(* IEC 61131-3 sources: daoli-st-library/DL_Device (part 19) *)

(* ---- FB_DL_DieCastCycleSupervise.st ---- *)
(*==============================================================================
  Component : FB_DL_DieCastCycleSupervise
  Category  : DL_Device
  Type      : FB
  Complexity: C4
  VERSION   : v1.0.0
  功能      : 压铸单循环监控与三级异常分级停机（黄记录 / 红判废 / 黑停机）
  开源溯源  : 道莅原创 clean-room 自研（无外部代码引用）｜License: MIT
  边界条件  : ① 压射曲线四点监控：慢速终点位置偏差（eSlowEndDev）、快射峰值速度（eFastVelLow）、
                 增压建立时间（eBuildSlow）、保压压力（eHoldLow）；四点各自独立判据与独立成因，
                 分级动作经 ApplyDefect 单点施加，禁共用枚举成员（R190）。
              ② 分级语义（写进契约）：黄 = 记录成因、本模继续；红 = 置 _bRejectMark 判废并单拍告警，
                 机械流程仍走到 eDone 才结算（废件必须被顶出取走，不得停在模内）；
                 黑 = 立即停机（超压 / 信号非有限 / 急停 / 安全门开），等 bReset 复位。
              ③ 判据限值配比约束（R100）：fSlowEndWarnMm ≤ fSlowEndTolMm、fFastVelWarnMps ≥ fFastVelMinMps、
                 fBuildWarnS ≤ fBuildMaxS、fHoldWarnMpa ≥ fHoldMinMpa；违反即组态非法（E2 黑前哨）。
              ④ 默认引脚组合自证（R114）：过程握手类（bClampClosed / bClampOpened / bEjectDone /
                 bPartTaken / bSprayDone / bRejectAck）默认 FALSE，默认组合无法推进任何相；使能类
                 （bEStopHealthy / bGuardClosed）默认 TRUE 与 bEnable 同族，断线由硬件安全回路保证。
              ⑤ 复位作用域（R311）：bReset 沿清 E2/E3 锁存 + 判废标记 + 分级 + 曲线锁存；bStop 只清 E2 与相位。
  状态机    : eIdle 待机 / eClampClose 合模 / eShotSlow 慢压射 / eShotFast 快压射 / eIntensify 增压 /
              eHold 保压 / eClampOpen 开模 / eEject 顶出 / eTakeOut 取件 / eSpray 喷涂 / eDone 结算拍 /
              eFault 停机待复位(E2) / eSafeStop 安全断能(E3)
  自检      : R1 零 GVL ｜ R2 零物理地址 ｜ R3 纯 IEC 61131-3 ｜ R4 非有限自反判 + 除法先判分母 ｜
              R6 CASE 含 ELSE ｜ R7 九 TON 两沿段 0 无条件刷新 ｜ R10 仅标准转换函数 ｜ R14 无属性件
==============================================================================*)
TYPE E_DL_DcsPhase :
(
    eIdle       := 0,   (* 待机：等启动沿 / Idle, waiting for start edge *)
    eClampClose := 10,  (* 合模：等合模到位 / Clamp closing *)
    eShotSlow   := 20,  (* 慢压射：到慢速终点 / Slow shot *)
    eShotFast   := 30,  (* 快压射：到快射终点 / Fast shot *)
    eIntensify  := 40,  (* 增压：建压到门限 / Intensification *)
    eHold       := 50,  (* 保压：保压到时 / Pressure hold *)
    eClampOpen  := 60,  (* 开模：等开模到位 / Clamp opening *)
    eEject      := 70,  (* 顶出：等顶出到位 / Ejecting *)
    eTakeOut    := 80,  (* 取件：等取件完成 / Take-out *)
    eSpray      := 90,  (* 喷涂：等喷涂完成 / Spraying *)
    eDone       := 100, (* 结算拍：模次与良率统计 / Settlement, one-scan *)
    eFault      := 120, (* 停机待复位（E2）/ Stop awaiting reset, E2 *)
    eSafeStop   := 130  (* 安全侧断能（E3）/ Safety energy cut, E3 *)
);
END_TYPE
TYPE E_DL_DcsCause :
(
    eNone       := 0,   (* 无异常 / No anomaly *)
    eSlowEndDev := 1,   (* 慢速终点位置偏差超限（红）/ Slow-shot end position deviation *)
    eFastVelLow := 2,   (* 快射速度偏低（黄或红）/ Fast-shot velocity low *)
    eBuildSlow  := 3,   (* 增压建立时间超限（黄或红）/ Intensification build too slow *)
    eHoldLow    := 4,   (* 保压压力偏低（黄或红）/ Hold pressure low *)
    ePressOver  := 5,   (* 压力超上限（黑）/ Over-pressure, black *)
    eSigBad     := 6,   (* 压力或位置信号非有限（黑）/ Non-finite signal, black *)
    eEStopOpen  := 7,   (* 急停回路断开（黑）/ E-stop open, black *)
    eGuardOpen  := 8,   (* 安全门未闭合（黑）/ Guard door open, black *)
    eClampTmo   := 9,   (* 合模或开模超时（黑）/ Clamp timeout, black *)
    eShotTmo    := 10,  (* 压射超时（黑）/ Shot timeout, black *)
    eBuildTmo   := 11,  (* 增压超时（黑）/ Intensify timeout, black *)
    eFastTmo    := 12,  (* 快射超时（黑）/ Fast-shot timeout, black *)
    eEjectTmo   := 13,  (* 顶出超时（黑）/ Eject timeout, black *)
    eTakeTmo    := 14,  (* 取件超时（黑）/ Take-out timeout, black *)
    eSprayTmo   := 15,  (* 喷涂超时（黑）/ Spray timeout, black *)
    eCfgBad     := 16,  (* 组态非法（E2）/ Illegal configuration, E2 *)
    ePhaseBad   := 17   (* 非法相位兜底（E2）/ Illegal phase fallback, E2 *)
);
END_TYPE
TYPE E_DL_DcsGrade :
(
    eOk     := 0,       (* 无异常：本模继续 / OK, continue *)
    eYellow := 1,       (* 黄：记录并继续，不置 bError / Yellow, recorded only *)
    eRed    := 2,       (* 红：本模判废并告警 / Red, part rejected with alarm *)
    eBlack  := 3        (* 黑：立即停机 / Black, immediate stop *)
);
END_TYPE

FUNCTION_BLOCK FB_DL_DieCastCycleSupervise
VAR_INPUT
    bStart          : BOOL := FALSE;    (* 启动沿（eIdle 入 eClampClose） [-] / Start rising edge *)
    bStop           : BOOL := FALSE;    (* 中止：回 eIdle 并清 E2 锁存 [-] / Abort, clears E2 only *)
    bReset          : BOOL := FALSE;    (* 复位沿：清全部锁存 + 曲线锁存（R311） [-] / Reset edge *)
    bRejectAck      : BOOL := FALSE;    (* 废模确认（只清告警标记，不推进相） [-] / Reject acknowledge *)
    bClampClosed    : BOOL := FALSE;    (* 合模到位（默认 FALSE 禁跳步） [-] / Clamp closed *)
    bClampOpened    : BOOL := FALSE;    (* 开模到位（默认 FALSE 禁跳步） [-] / Clamp opened *)
    bEjectDone      : BOOL := FALSE;    (* 顶出到位（默认 FALSE 禁跳步） [-] / Eject done *)
    bPartTaken      : BOOL := FALSE;    (* 取件完成（默认 FALSE 禁跳步） [-] / Part taken *)
    bSprayDone      : BOOL := FALSE;    (* 喷涂完成（默认 FALSE 禁跳步） [-] / Spray done *)
    bGuardClosed    : BOOL := TRUE;     (* 安全门闭合（使能类引脚，默认 TRUE） [-] / Guard door closed *)
    bEStopHealthy   : BOOL := TRUE;     (* 急停回路正常（使能类引脚，默认 TRUE） [-] / E-stop healthy *)
    fShotPosMm      : LREAL := 0.0;     (* 冲头实时位置（0 = 起始位） [mm] / Shot position [mm] *)
    fShotVelMps     : LREAL := 0.0;     (* 冲头实时速度 [m/s] / Shot velocity [m/s] *)
    fHoldPressMpa   : LREAL := 0.0;     (* 压射缸压力实测 [MPa] / Shot pressure [MPa] *)
    fSlowEndSetMm   : LREAL := 250.0;   (* 慢速终点设定位置，域 > 0 [mm] / Slow-end setpoint [mm] *)
    fShotEndMm      : LREAL := 320.0;   (* 快射终点位置，域 > fSlowEndSetMm [mm] / Fast-shot end [mm] *)
    fSlowEndWarnMm  : LREAL := 10.0;    (* 慢速终点偏差预警限（黄），域 >= 0 [mm] / Slow-end warn limit [mm] *)
    fSlowEndTolMm   : LREAL := 25.0;    (* 慢速终点偏差硬限（红），域 > 0 [mm] / Slow-end hard limit [mm] *)
    fFastVelMinMps  : LREAL := 2.5;     (* 快射速度硬下限（红），域 > 0 [m/s] / Fast velocity hard min [m/s] *)
    fFastVelWarnMps : LREAL := 3.0;     (* 快射速度预警下限（黄），域 > 0 [m/s] / Fast velocity warn min [m/s] *)
    fIntensifyMpa   : LREAL := 18.0;    (* 增压建立压力门限，域 > 0 [MPa] / Build threshold [MPa] *)
    fBuildWarnS     : LREAL := 0.08;    (* 增压建立时间预警限（黄），域 >= 0 [s] / Build warn limit [s] *)
    fBuildMaxS      : LREAL := 0.15;    (* 增压建立时间硬限（红），域 > 0 [s] / Build hard limit [s] *)
    fHoldMinMpa     : LREAL := 12.0;    (* 保压压力硬下限（红），域 > 0 [MPa] / Hold pressure hard min [MPa] *)
    fHoldWarnMpa    : LREAL := 14.0;    (* 保压压力预警下限（黄），域 > 0 [MPa] / Hold pressure warn min [MPa] *)
    fPressOverMpa   : LREAL := 30.0;    (* 压力超上限（黑断能），域 > 0 [MPa] / Over-pressure limit [MPa] *)
    atPhaseTmo      : ARRAY[0..8] OF TIME := [T#10S, T#5S, T#5S, T#5S, T#30S, T#10S, T#10S, T#15S, T#15S];   (* 超时窗 [ms]，下标 0..8 = 合模/慢射/快射/增压/保压/开模/顶出/取件/喷涂 / Phase windows [ms] *)
    fCycleSec       : LREAL := 0.0;     (* 扫描周期（<=0 用缺省 0.01s） [s] / Scan cycle [s] *)
END_VAR
VAR_OUTPUT
    eState          : E_DL_DcsPhase;    (* 当前相（HMI 诊断） [-] / Present phase *)
    eCause          : E_DL_DcsCause;    (* 成因（锁存回放，R189） [-] / Latched cause playback *)
    eGrade          : E_DL_DcsGrade;    (* 本模判据分级（黄/红/黑）；组态 E2 不改分级、由 bError 表达 [-] / Criterion grade, E2 config fault expressed by bError *)
    bError          : BOOL;             (* 故障标志（仅黑与 E2 置位，黄/红不置） [-] / Error flag *)
    bSafeCut        : BOOL;             (* 安全侧断能指令（黑常 TRUE 至复位） [-] / Safety energy cut *)
    bReject         : BOOL;             (* 本模判废标告警（红级置位，结算或确认后清） [-] / Reject alarm *)
    bDone           : BOOL;             (* 单拍结算脉冲 [-] / One-scan done pulse *)
    bShotActive     : BOOL;             (* 压射段指示（供 IO 层驱动压射阀） [-] / Shot indicator *)
    nShotCount      : UDINT;            (* 累计模次（饱和） [模] / Shot count, saturating *)
    nGoodCount      : UDINT;            (* 累计良品（饱和） [模] / Good part count *)
    fYieldPct       : LREAL;            (* 良率（无模次输出 0） [%] / Yield [%] *)
    fSlowEndLastMm  : LREAL;            (* 最近一模慢速终点实测 [mm] / Last slow-end position [mm] *)
    fFastVelLastMps : LREAL;            (* 最近一模快射峰值速度 [m/s] / Last peak velocity [m/s] *)
    fBuildLastS     : LREAL;            (* 最近一模增压建立时间 [s] / Last build time [s] *)
    fHoldLastMpa    : LREAL;            (* 最近一模保压压力 [MPa] / Last hold pressure [MPa] *)
END_VAR
VAR
    _ePhase      : E_DL_DcsPhase := E_DL_DcsPhase.eIdle;     (* 内部相（CASE 唯一写入目标） [-] / Internal phase *)
    _eCause      : E_DL_DcsCause := E_DL_DcsCause.eNone;     (* 成因锁存量 [-] / Latched cause *)
    _eGrade      : E_DL_DcsGrade := E_DL_DcsGrade.eOk;       (* 本模分级锁存量 [-] / Latched grade *)
    _bFault      : BOOL := FALSE;       (* E2 锁存位（解除 = bReset 沿或 bStop） [-] / E2 latch *)
    _bSafeLatch  : BOOL := FALSE;       (* E3 锁存位（解除 = bReset 沿且安全恢复） [-] / E3 latch *)
    _bFaultReq   : BOOL := FALSE;       (* 单拍 E2 请求（段 1 预清，段 6 落地） [-] / One-scan E2 request *)
    _bSafeReq    : BOOL := FALSE;       (* 单拍 E3 请求（段 1 预清，段 6 落地） [-] / One-scan E3 request *)
    _bDonePulse  : BOOL := FALSE;       (* 单拍结算标志（段 1 预清） [-] / One-scan done flag *)
    _bRejectMark : BOOL := FALSE;       (* 本模判废标记（红级置位，结算清零） [-] / Reject mark for this shot *)
    _bPressBad   : BOOL := FALSE;       (* 压力信号非有限当拍量 [-] / Pressure non-finite *)
    _bPosBad     : BOOL := FALSE;       (* 位置信号非有限当拍量 [-] / Position non-finite *)
    _bVelBad     : BOOL := FALSE;       (* 速度信号非有限当拍量 [-] / Velocity non-finite *)
    _bBuilt      : BOOL := FALSE;       (* 增压已建立（当拍判据） [-] / Intensification built *)
    _bCfgBad     : BOOL := FALSE;       (* 组态非法当拍量 [-] / Configuration bad *)
    _nIdxChk     : INT := 0;            (* 相窗遍历索引（循环变量） [-] / Loop index *)
    _fCy         : LREAL := 0.0;        (* 当拍有效周期 [s] / Effective cycle *)
    _fVelPeak    : LREAL := 0.0;        (* 快射峰值速度（入快射相清零） [m/s] / Fast-shot peak [m/s] *)
    _fBuildS     : LREAL := 0.0;        (* 增压建立时间累加（入增压相清零） [s] / Build time accumulator [s] *)
    _fSlowEndMm  : LREAL := 0.0;        (* 慢速终点位置锁存 [mm] / Slow-end position latch *)
    _fHoldMpa    : LREAL := 0.0;        (* 保压压力锁存 [MPa] / Hold pressure latch *)
    _nShot       : UDINT := 0;          (* 模次累计锁存（饱和） [模] / Shot count latch *)
    _nGood       : UDINT := 0;          (* 良品累计锁存（饱和） [模] / Good count latch *)
    tonClampClose: TON;                 (* 合模超时（段 0 无条件调用） / Clamp-close timeout *)
    tonShotSlow  : TON;                 (* 慢压射超时 / Slow-shot timeout *)
    tonShotFast  : TON;                 (* 快压射超时 / Fast-shot timeout *)
    tonIntensify : TON;                 (* 增压超时 / Intensify timeout *)
    tonHold      : TON;                 (* 保压计时与超时 / Hold timer *)
    tonClampOpen : TON;                 (* 开模超时 / Clamp-open timeout *)
    tonEject     : TON;                 (* 顶出超时 / Eject timeout *)
    tonTakeOut   : TON;                 (* 取件超时 / Take-out timeout *)
    tonSpray     : TON;                 (* 喷涂超时 / Spray timeout *)
    rtStart      : R_TRIG;              (* 启动沿（段 0 无条件调用） / Start edge *)
    rtReset      : R_TRIG;              (* 复位沿（段 0 无条件调用） / Reset edge *)
END_VAR
VAR CONSTANT
    DL_DCS_CYDEF   : LREAL := 0.01;         (* 缺省扫描周期 [s] / Default scan cycle [s] *)
    DL_DCS_CNTMAX  : UDINT := 4294967295;   (* 模次与良品计数饱和上限 [模] / Count ceiling *)
    DL_DCS_PCTOP   : LREAL := 100.0;        (* 良率百分比满量程 [%] / Yield full scale [%] *)
END_VAR

(*-----------------------------------------------------------------------------
  方法 GradeFault：单点判据分级（纯分类，不修改任何 FB 状态）
  契约：fValue 为「按变差方向已归一」的判据量（偏差取绝对值后传入）；
        bLowerWorse = TRUE 表示低于限值变差，FALSE 表示高于限值变差；
        fWarnLimit 必须落在「正常侧」，fHardLimit 落在「变差侧」（配比由组态闸保证）。
        非有限实测（NaN 自反 / Inf 差值自减）一律返回 eBlack：信号失效必须停机。
-----------------------------------------------------------------------------*)
METHOD PUBLIC GradeFault : E_DL_DcsGrade
VAR_INPUT
    fValue      : LREAL := 0.0;     (* 判据实测值（已按方向归一） [工程单位] / Measured criterion *)
    fWarnLimit  : LREAL := 0.0;     (* 预警限（黄级） [工程单位] / Warning limit *)
    fHardLimit  : LREAL := 0.0;     (* 硬限（红级） [工程单位] / Hard limit *)
    bLowerWorse : BOOL := FALSE;    (* TRUE = 低于限值变差 [-] / Lower is worse when TRUE *)
END_VAR

GradeFault := E_DL_DcsGrade.eOk;    (* 预置：无异常 / Preset OK *)
IF (fValue <> fValue) OR ((fValue - fValue) <> (fValue - fValue)) THEN
    GradeFault := E_DL_DcsGrade.eBlack;     (* 非有限 -> 黑级停机 / Non-finite, black *)
    RETURN;
END_IF
IF bLowerWorse THEN
    IF fValue < fHardLimit THEN
        GradeFault := E_DL_DcsGrade.eRed;   (* 低于硬限 -> 红 / Below hard limit *)
    ELSIF fValue < fWarnLimit THEN
        GradeFault := E_DL_DcsGrade.eYellow;(* 低于预警限 -> 黄 / Below warn limit *)
    END_IF
ELSE
    IF fValue > fHardLimit THEN
        GradeFault := E_DL_DcsGrade.eRed;   (* 高于硬限 -> 红 / Above hard limit *)
    ELSIF fValue > fWarnLimit THEN
        GradeFault := E_DL_DcsGrade.eYellow;(* 高于预警限 -> 黄 / Above warn limit *)
    END_IF
END_IF
END_METHOD

(*-----------------------------------------------------------------------------
  方法 ApplyDefect：分级动作单点施加（唯一写入 _eGrade / _bRejectMark / _bSafeReq 的位置）
  契约：eOk 不写任何量；eBlack 只请求 E3（由段 6 落地并迁相）；eRed 置判废标记与告警；
        eYellow 只在尚未升级到红/黑时记录。分级只升不降（本模内单调）。
-----------------------------------------------------------------------------*)
METHOD PRIVATE ApplyDefect
VAR_INPUT
    xGrade : E_DL_DcsGrade := E_DL_DcsGrade.eOk;    (* 分级结果 [-] / Grade result *)
    xCause : E_DL_DcsCause := E_DL_DcsCause.eNone;  (* 归因（各判据点独立传入） [-] / Cause per point *)
END_VAR

IF xGrade = E_DL_DcsGrade.eOk THEN
    RETURN;                                     (* 无异常：不写任何量 / Nothing to apply *)
END_IF
_eCause := xCause;                              (* 归因：调用点唯一指定 / Cause assigned by caller *)
IF xGrade = E_DL_DcsGrade.eBlack THEN
    _bSafeReq := TRUE;                          (* 黑级：请求 E3 断能 / Black: request E3 *)
ELSIF xGrade = E_DL_DcsGrade.eRed THEN
    IF _eGrade <> E_DL_DcsGrade.eBlack THEN
        _eGrade := E_DL_DcsGrade.eRed;          (* 红级：判废（黑级不被降级）/ Red, never downgrade black *)
    END_IF
    _bRejectMark := TRUE;                       (* 本模判废标记 / Reject mark *)
ELSIF _eGrade = E_DL_DcsGrade.eOk THEN
    _eGrade := E_DL_DcsGrade.eYellow;           (* 黄级：仅当尚未升级时记录 / Yellow only if still OK *)
END_IF
END_METHOD

(*-----------------------------------------------------------------------------
  方法 ResetCycle：本模曲线锁存与分级复位（不清累计模次与良品数）
  契约：返回 TRUE 表示复位执行；作用于分级、判废标记与四点曲线锁存；
        累计计数（_nShot / _nGood）属生产资料，只能由 bReset 沿清除，本方法不动。
-----------------------------------------------------------------------------*)
METHOD PUBLIC ResetCycle : BOOL
ResetCycle := FALSE;                            (* 预置 / Preset *)
_eGrade := E_DL_DcsGrade.eOk;                   (* 清分级 / Clear grade *)
_eCause := E_DL_DcsCause.eNone;                 (* 清成因 / Clear cause *)
_bRejectMark := FALSE;                          (* 清判废标记 / Clear reject mark *)
_fVelPeak := 0.0;                               (* 清快射峰值 / Clear peak *)
_fBuildS := 0.0;                                (* 清建立时间 / Clear build time *)
_fSlowEndMm := 0.0;                             (* 清慢速终点锁存 / Clear slow-end latch *)
_fHoldMpa := 0.0;                               (* 清保压压力锁存 / Clear hold latch *)
ResetCycle := TRUE;                             (* 复位已执行 / Reset performed *)
END_METHOD

(* —— 段 0：三测量量非有限判定 + 组态闸 + 周期派生 + 峰值与建压跟踪 + 九 TON 两沿无条件刷新（R7） —— *)
_bPressBad := (fHoldPressMpa <> fHoldPressMpa)
           OR ((fHoldPressMpa - fHoldPressMpa) <> (fHoldPressMpa - fHoldPressMpa));   (* NaN 自反 + Inf 差值 / NaN and Inf *)
_bPosBad := (fShotPosMm <> fShotPosMm)
         OR ((fShotPosMm - fShotPosMm) <> (fShotPosMm - fShotPosMm));
_bVelBad := (fShotVelMps <> fShotVelMps)
         OR ((fShotVelMps - fShotVelMps) <> (fShotVelMps - fShotVelMps));
_bCfgBad := (fSlowEndSetMm <= 0.0) OR (fShotEndMm <= fSlowEndSetMm) OR (fSlowEndTolMm <= 0.0) OR (fSlowEndWarnMm < 0.0)
         OR (fSlowEndWarnMm > fSlowEndTolMm)                       (* 限值配比① / Ratio 1 *)
         OR (fFastVelMinMps <= 0.0) OR (fFastVelWarnMps <= 0.0)
         OR (fFastVelWarnMps < fFastVelMinMps)                     (* 限值配比② / Ratio 2 *)
         OR (fIntensifyMpa <= 0.0) OR (fBuildMaxS <= 0.0) OR (fBuildWarnS < 0.0)
         OR (fBuildWarnS > fBuildMaxS)                             (* 限值配比③ / Ratio 3 *)
         OR (fHoldMinMpa <= 0.0) OR (fHoldWarnMpa <= 0.0)
         OR (fHoldWarnMpa < fHoldMinMpa)                           (* 限值配比④ / Ratio 4 *)
         OR (fPressOverMpa <= fHoldWarnMpa);                       (* 超压限须高于保压下限 / Over limit above hold *)
FOR _nIdxChk := 0 TO 8 DO
    IF atPhaseTmo[_nIdxChk] <= T#0S THEN
        _bCfgBad := TRUE;                                          (* 任一相窗非正 -> 组态非法 / Non-positive window *)
    END_IF
END_FOR
IF fCycleSec > 0.0 THEN
    _fCy := fCycleSec;                                             (* 组态周期有效 / Configured cycle *)
ELSE
    _fCy := DL_DCS_CYDEF;                                          (* 周期缺省兜底 / Default cycle *)
END_IF
_bBuilt := (_ePhase = E_DL_DcsPhase.eIntensify) AND (NOT _bPressBad) AND (fHoldPressMpa >= fIntensifyMpa);
IF (_ePhase = E_DL_DcsPhase.eIntensify) AND (NOT _bBuilt) THEN
    _fBuildS := _fBuildS + _fCy;                                   (* 增压建立时间累加 [s] / Build time accumulation *)
END_IF
IF (_ePhase = E_DL_DcsPhase.eShotFast) AND (NOT _bVelBad) THEN
    IF fShotVelMps > _fVelPeak THEN
        _fVelPeak := fShotVelMps;                                  (* 快射峰值跟踪 / Peak tracking *)
    END_IF
END_IF
rtStart(CLK := bStart);                                            (* 启动沿，每拍必调 / Start edge every scan *)
rtReset(CLK := bReset);                                            (* 复位沿，每拍必调 / Reset edge every scan *)
tonClampClose(IN := (_ePhase = E_DL_DcsPhase.eClampClose), PT := atPhaseTmo[0]);   (* 合模窗 / Clamp window *)
tonShotSlow(IN := (_ePhase = E_DL_DcsPhase.eShotSlow), PT := atPhaseTmo[1]);       (* 慢射窗 / Slow shot window *)
tonShotFast(IN := (_ePhase = E_DL_DcsPhase.eShotFast), PT := atPhaseTmo[2]);       (* 快射窗 / Fast shot window *)
tonIntensify(IN := (_ePhase = E_DL_DcsPhase.eIntensify), PT := atPhaseTmo[3]);     (* 增压窗 / Intensify window *)
tonHold(IN := (_ePhase = E_DL_DcsPhase.eHold), PT := atPhaseTmo[4]);               (* 保压窗 / Hold window *)
tonClampOpen(IN := (_ePhase = E_DL_DcsPhase.eClampOpen), PT := atPhaseTmo[5]);     (* 开模窗 / Open window *)
tonEject(IN := (_ePhase = E_DL_DcsPhase.eEject), PT := atPhaseTmo[6]);             (* 顶出窗 / Eject window *)
tonTakeOut(IN := (_ePhase = E_DL_DcsPhase.eTakeOut), PT := atPhaseTmo[7]);         (* 取件窗 / Take-out window *)
tonSpray(IN := (_ePhase = E_DL_DcsPhase.eSpray), PT := atPhaseTmo[8]);             (* 喷涂窗 / Spray window *)

(* —— 段 1：单拍量预清零（不含锁存/计数/曲线量，R107） —— *)
_bFaultReq := FALSE;                                               (* E2 请求预清 / E2 request preset *)
_bSafeReq := FALSE;                                                (* E3 请求预清 / E3 request preset *)
_bDonePulse := FALSE;                                              (* 结算标志预清 / Done preset *)
bError := FALSE;                                                   (* 故障标志预清（出口汇总）/ Error preset *)

(* —— 段 2：黑级安全侧（急停 / 安全门 / 超压 / 压力与位置信号非有限）——最高优先级 —— *)
IF (NOT bEStopHealthy) OR (NOT bGuardClosed) THEN
    IF NOT _bSafeLatch THEN
        _bSafeReq := TRUE;                                         (* 落地于段 6 / Landed in segment 6 *)
        IF NOT bEStopHealthy THEN
            _eCause := E_DL_DcsCause.eEStopOpen;                   (* 归因：急停断开 / Cause: E-stop *)
        ELSE
            _eCause := E_DL_DcsCause.eGuardOpen;                   (* 归因：安全门开 / Cause: guard *)
        END_IF
    END_IF
ELSIF _bPressBad OR _bPosBad THEN
    IF NOT _bSafeLatch THEN
        _bSafeReq := TRUE;
        _eCause := E_DL_DcsCause.eSigBad;                          (* 归因：信号非有限 / Cause: non-finite *)
    END_IF
ELSIF (NOT _bPressBad) AND (fHoldPressMpa > fPressOverMpa) THEN
    IF NOT _bSafeLatch THEN
        _bSafeReq := TRUE;
        _eCause := E_DL_DcsCause.ePressOver;                       (* 归因：超压 / Cause: over-pressure *)
    END_IF
END_IF

(* —— 段 3：组态闸入 E2（黑级优先，安全相内不重复置因） —— *)
IF _bCfgBad AND (NOT _bSafeLatch) AND (NOT _bFault) THEN
    _bFaultReq := TRUE;                                            (* 落地于段 6 / Landed in segment 6 *)
    _eCause := E_DL_DcsCause.eCfgBad;                              (* 归因：组态非法 / Cause: config *)
END_IF

(* —— 段 4：迁出链（复位沿 > 中止 > 废模确认；作用域逐项声明 R311） —— *)
IF rtReset.Q THEN
    _bFault := FALSE;                                              (* 作用域①：清 E2 锁存 / Clear E2 *)
    IF NOT ((NOT bEStopHealthy) OR (NOT bGuardClosed) OR _bPressBad OR _bPosBad
            OR ((NOT _bPressBad) AND (fHoldPressMpa > fPressOverMpa))) THEN
        _bSafeLatch := FALSE;                                      (* 作用域②：安全恢复才清 E3 / Clear E3 only if safe *)
    END_IF
    _eCause := E_DL_DcsCause.eNone;                                (* 作用域③：清成因与分级 / Clear cause and grade *)
    _eGrade := E_DL_DcsGrade.eOk;
    _bRejectMark := FALSE;                                         (* 作用域④：清判废标记 / Clear reject mark *)
    _fVelPeak := 0.0;                                              (* 作用域⑤：清曲线锁存 / Clear curve latches *)
    _fBuildS := 0.0;
    _nShot := 0;                                                   (* 作用域⑥：清模次与良品（生产资料复位）/ Clear counters *)
    _nGood := 0;
    IF NOT _bSafeLatch THEN
        IF (_ePhase = E_DL_DcsPhase.eFault) OR (_ePhase = E_DL_DcsPhase.eSafeStop) THEN
            _ePhase := E_DL_DcsPhase.eIdle;                        (* 作用域⑦：故障相迁回待机 / Back to idle *)
        END_IF
    END_IF
ELSIF bStop AND (_ePhase <> E_DL_DcsPhase.eIdle) AND (_ePhase <> E_DL_DcsPhase.eSafeStop) THEN
    IF _ePhase = E_DL_DcsPhase.eFault THEN
        _bFault := FALSE;                                          (* 中止清 E2（E3 只由复位清）/ Abort clears E2 only *)
        _eCause := E_DL_DcsCause.eNone;
        _eGrade := E_DL_DcsGrade.eOk;
    END_IF
    _ePhase := E_DL_DcsPhase.eIdle;                                (* 回待机 / Back to idle *)
ELSIF bRejectAck THEN
    _bRejectMark := FALSE;                                         (* 废模确认只清告警标记 / Ack clears alarm only *)
END_IF

(* —— 段 5：主状态机（四点曲线判据在相迁移点判定，动作经 ApplyDefect 单点施加） —— *)
CASE _ePhase OF
E_DL_DcsPhase.eIdle:
    IF rtStart.Q AND (NOT _bFault) AND (NOT _bSafeLatch) THEN
        _eGrade := E_DL_DcsGrade.eOk;                              (* 新模起算 / New shot *)
        _eCause := E_DL_DcsCause.eNone;
        _bRejectMark := FALSE;
        _ePhase := E_DL_DcsPhase.eClampClose;                      (* 入合模相 / To clamp close *)
    END_IF
E_DL_DcsPhase.eClampClose:
    IF bClampClosed THEN
        _ePhase := E_DL_DcsPhase.eShotSlow;                        (* 合模到位 -> 慢压射 / Clamped, slow shot *)
    ELSIF tonClampClose.Q THEN
        _eCause := E_DL_DcsCause.eClampTmo;                        (* 归因：合模超时 / Cause: clamp timeout *)
        _bSafeReq := TRUE;
    END_IF
E_DL_DcsPhase.eShotSlow:
    IF (NOT _bPosBad) AND (fShotPosMm >= fSlowEndSetMm) THEN
        _fSlowEndMm := fShotPosMm;                                 (* 慢速终点锁存 / Latch slow end *)
        ApplyDefect(GradeFault(ABS(_fSlowEndMm - fSlowEndSetMm), fSlowEndWarnMm, fSlowEndTolMm, FALSE),
                    E_DL_DcsCause.eSlowEndDev);                    (* 判据点①：慢速终点偏差 / Point 1 *)
        _fVelPeak := 0.0;                                          (* 快射峰值起算 / Peak restart *)
        _ePhase := E_DL_DcsPhase.eShotFast;                        (* 入快压射相 / To fast shot *)
    ELSIF tonShotSlow.Q THEN
        _eCause := E_DL_DcsCause.eShotTmo;                         (* 归因：慢射超时 / Cause: slow-shot timeout *)
        _bSafeReq := TRUE;
    END_IF
E_DL_DcsPhase.eShotFast:
    IF (NOT _bPosBad) AND (fShotPosMm >= fShotEndMm) THEN
        ApplyDefect(GradeFault(_fVelPeak, fFastVelWarnMps, fFastVelMinMps, TRUE),
                    E_DL_DcsCause.eFastVelLow);                    (* 判据点②：快射峰值速度 / Point 2 *)
        _fBuildS := 0.0;                                           (* 建压计时起算 / Build restart *)
        _ePhase := E_DL_DcsPhase.eIntensify;                       (* 入增压相 / To intensify *)
    ELSIF tonShotFast.Q THEN
        _eCause := E_DL_DcsCause.eFastTmo;                         (* 归因：快射超时 / Cause: fast-shot timeout *)
        _bSafeReq := TRUE;
    END_IF
E_DL_DcsPhase.eIntensify:
    IF _bBuilt THEN
        ApplyDefect(GradeFault(_fBuildS, fBuildWarnS, fBuildMaxS, FALSE),
                    E_DL_DcsCause.eBuildSlow);                     (* 判据点③：增压建立时间 / Point 3 *)
        _ePhase := E_DL_DcsPhase.eHold;                            (* 建压完成 -> 保压 / Built, hold *)
    ELSIF tonIntensify.Q THEN
        _eCause := E_DL_DcsCause.eBuildTmo;                        (* 归因：增压超时 / Cause: build timeout *)
        _bSafeReq := TRUE;
    END_IF
E_DL_DcsPhase.eHold:
    IF tonHold.Q THEN
        _fHoldMpa := fHoldPressMpa;                                (* 保压压力锁存 / Latch hold pressure *)
        ApplyDefect(GradeFault(_fHoldMpa, fHoldWarnMpa, fHoldMinMpa, TRUE),
                    E_DL_DcsCause.eHoldLow);                       (* 判据点④：保压压力 / Point 4 *)
        _ePhase := E_DL_DcsPhase.eClampOpen;                       (* 保压到时 -> 开模 / Hold done, open *)
    END_IF
E_DL_DcsPhase.eClampOpen:
    IF bClampOpened THEN
        _ePhase := E_DL_DcsPhase.eEject;                           (* 开模到位 -> 顶出 / Opened, eject *)
    ELSIF tonClampOpen.Q THEN
        _eCause := E_DL_DcsCause.eClampTmo;                        (* 归因：开模超时 / Cause: open timeout *)
        _bSafeReq := TRUE;
    END_IF
E_DL_DcsPhase.eEject:
    IF bEjectDone THEN
        _ePhase := E_DL_DcsPhase.eTakeOut;                         (* 顶出到位 -> 取件 / Ejected, take out *)
    ELSIF tonEject.Q THEN
        _eCause := E_DL_DcsCause.eEjectTmo;                        (* 归因：顶出超时 / Cause: eject timeout *)
        _bSafeReq := TRUE;
    END_IF
E_DL_DcsPhase.eTakeOut:
    IF bPartTaken THEN
        _ePhase := E_DL_DcsPhase.eSpray;                           (* 取件完成 -> 喷涂 / Taken, spray *)
    ELSIF tonTakeOut.Q THEN
        _eCause := E_DL_DcsCause.eTakeTmo;                         (* 归因：取件超时 / Cause: take-out timeout *)
        _bSafeReq := TRUE;
    END_IF
E_DL_DcsPhase.eSpray:
    IF bSprayDone THEN
        _ePhase := E_DL_DcsPhase.eDone;                            (* 喷涂完成 -> 结算 / Sprayed, settle *)
    ELSIF tonSpray.Q THEN
        _eCause := E_DL_DcsCause.eSprayTmo;                        (* 归因：喷涂超时 / Cause: spray timeout *)
        _bSafeReq := TRUE;
    END_IF
E_DL_DcsPhase.eDone:
    _bDonePulse := TRUE;                                           (* 单拍结算（段 1 预清）/ One-scan done *)
    IF _nShot < DL_DCS_CNTMAX THEN
        _nShot := _nShot + 1;                                      (* 模次推进（容量载体判上限）/ Saturating shot count *)
    END_IF
    IF (NOT _bRejectMark) AND (_nGood < DL_DCS_CNTMAX) THEN
        _nGood := _nGood + 1;                                      (* 良品推进（判废模不计良）/ Saturating good count *)
    END_IF
    _ePhase := E_DL_DcsPhase.eIdle;                                (* 回待机迎下一模 / Back to idle *)
E_DL_DcsPhase.eFault:
    bError := TRUE;                                                (* 故障相驻留（锁存回放）/ Fault residency *)
E_DL_DcsPhase.eSafeStop:
    bError := TRUE;                                                (* 安全相驻留（锁存回放）/ Safety residency *)
ELSE
    _eCause := E_DL_DcsCause.ePhaseBad;                            (* 非法相位兜底 / Illegal phase fallback *)
    _bFaultReq := TRUE;                                            (* 由段 6 落地 / Landed in segment 6 *)
END_CASE

(* —— 段 6：E2/E3 请求统一落地（分支内只写成因与请求，落地仅此一处，R187/R252） —— *)
IF _bSafeReq AND (NOT _bSafeLatch) THEN
    _bSafeLatch := TRUE;                                           (* E3 锁存（黑级）/ Latch E3 *)
    _eGrade := E_DL_DcsGrade.eBlack;                               (* 分级黑 / Grade black *)
    _ePhase := E_DL_DcsPhase.eSafeStop;                            (* 同步迁相 / Migrate *)
    bError := TRUE;                                                (* 故障标志同段置位（R45 配对）/ Error pairing *)
ELSIF _bFaultReq AND (NOT _bSafeLatch) THEN
    _bFault := TRUE;                                               (* E2 锁存 / Latch E2 *)
    _ePhase := E_DL_DcsPhase.eFault;                               (* 同步迁相（R252）/ Migrate *)
    bError := TRUE;                                                (* 故障标志同段置位（R45 配对）/ Error pairing *)
END_IF

(* —— 段 7：统一出口（电平量由 _ePhase 派生，计数与良率带零除守卫） —— *)
eState := _ePhase;                                                 (* 相出口 / Phase outlet *)
eCause := _eCause;                                                 (* 成因回放 / Cause playback *)
eGrade := _eGrade;                                                 (* 分级出口 / Grade outlet *)
bError := bError OR _bFault OR _bSafeLatch;                        (* 故障标志汇总（黄/红不置）/ Error summary *)
bSafeCut := _bSafeLatch;                                           (* 安全断能指令 / Safety energy cut *)
bReject := _bRejectMark;                                           (* 判废告警（红级）/ Reject alarm *)
bDone := _bDonePulse;                                              (* 单拍结算脉冲 / One-scan done *)
bShotActive := (_ePhase = E_DL_DcsPhase.eShotSlow) OR (_ePhase = E_DL_DcsPhase.eShotFast)
            OR (_ePhase = E_DL_DcsPhase.eIntensify);               (* 压射段指示 / Shot indicator *)
nShotCount := _nShot;                                              (* 模次出口 / Shot count outlet *)
nGoodCount := _nGood;                                              (* 良品出口 / Good count outlet *)
IF _nShot > 0 THEN
    fYieldPct := (UDINT_TO_LREAL(_nGood) / UDINT_TO_LREAL(_nShot)) * DL_DCS_PCTOP;   (* 良率（分母已判非零）/ Guarded yield *)
ELSE
    fYieldPct := 0.0;                                              (* 无模次输出 0 / No shot, zero *)
END_IF
fSlowEndLastMm := _fSlowEndMm;                                     (* 慢速终点出口 / Slow-end outlet *)
fFastVelLastMps := _fVelPeak;                                      (* 快射峰值出口 / Peak velocity outlet *)
fBuildLastS := _fBuildS;                                           (* 建立时间出口 / Build time outlet *)
fHoldLastMpa := _fHoldMpa;                                         (* 保压压力出口 / Hold pressure outlet *)
END_FUNCTION_BLOCK

(* ---- FB_DL_DieSprayReleaseSeq.st ---- *)
(*
  Component : FB_DL_DieSprayReleaseSeq
  Category  : DL_Device
  Type      : FB
  Complexity: C2
  VERSION   : v1.0.0
  功能      : 喷涂脱模剂时序控制：ENUM 七态（Idle/Open/Spray/Blow/Close/Done/Fault），按设定喷涂次数循环喷涂-吹扫，末次吹扫后关模。
  开源溯源  : 道莅原创 clean-room 自研（无外部代码引用）｜License: MIT
  边界条件  : ① 喷涂次数须 >= 1、四段时长均须非 0，否则拒绝启动并锁存故障码；
              ② 喷涂计数在喷涂段迁出拍单点累加，不在段内每拍累加；
              ③ 故障锁存唯一解除路径 = bReset 上升沿；eDone 撤销 bStart 回 eIdle。
*)

TYPE E_DL_SprayPhase :
(
    eIdle  := 0,    (* 空闲：等启动沿 / Idle waiting start edge *)
    eOpen  := 10,   (* 开模：开模动作 / Die opening *)
    eSpray := 20,   (* 喷涂：单次喷涂 / Single spray shot *)
    eBlow  := 30,   (* 吹扫：残液吹扫 / Air blow-off *)
    eClose := 40,   (* 关模：关模动作 / Die closing *)
    eDone  := 50,   (* 完成：驻留待撤销 / Done holding *)
    eFault := 90    (* 故障：锁存待复位 / Fault latched *)
);
END_TYPE

FUNCTION_BLOCK FB_DL_DieSprayReleaseSeq
VAR_INPUT
    bEnable   : BOOL;   (* 使能电平 [-] Enable level *)
    bReset    : BOOL;   (* 复位上升沿，清故障锁存 [-] Reset edge *)
    bStart    : BOOL;   (* 启动上升沿 [-] Start edge *)
    nSpraySet : INT;    (* 设定喷涂次数 [次] Spray shot count setpoint *)
    tOpen     : TIME;   (* 开模动作时长 [ms] Die opening duration *)
    tSpray    : TIME;   (* 单次喷涂时长 [ms] Spray shot duration *)
    tBlow     : TIME;   (* 吹扫时长 [ms] Air blow duration *)
    tClose    : TIME;   (* 关模动作时长 [ms] Die closing duration *)
END_VAR
VAR_OUTPUT
    bOpenCmd   : BOOL;               (* 开模指令 [-] Die open command *)
    bSprayCmd  : BOOL;               (* 喷涂指令 [-] Spray command *)
    bBlowCmd   : BOOL;               (* 吹扫指令 [-] Air blow command *)
    bCloseCmd  : BOOL;               (* 关模指令 [-] Die close command *)
    nSprayDone : INT;                (* 已完成喷涂次数 [次] Completed spray shots *)
    ePhase     : E_DL_SprayPhase;    (* 相位出口，段尾单点映射 [-] Phase outlet *)
    bError     : BOOL;               (* 故障锁存标志 [-] Fault latch flag *)
    uErrId     : UDINT;              (* 事件码，0 = 无事件 [-] Event code *)
END_VAR
VAR
    rtReset  : R_TRIG;   (* 复位沿实例，每拍无条件刷新 / Reset edge *)
    rtStart  : R_TRIG;   (* 启动沿实例，每拍无条件刷新 / Start edge *)
    tonOpen  : TON;      (* 开模动作计时（独立实例） / Open timer *)
    tonSpray : TON;      (* 喷涂计时（独立实例） / Spray timer *)
    tonBlow  : TON;      (* 吹扫计时（独立实例） / Blow timer *)
    tonClose : TON;      (* 关模动作计时（独立实例） / Close timer *)
    _ePhase  : E_DL_SprayPhase := E_DL_SprayPhase.eIdle;  (* 内部相位 / Internal phase *)
    _bFault  : BOOL;     (* 故障锁存位（锁存量） / Latched fault bit *)
    _uFault  : UDINT;    (* 故障码锁存（锁存量） / Latched fault code *)
    _bCfgBad : BOOL;     (* 组态非法当拍量 [-] Config illegal flag *)
END_VAR

(* —— 段 0｜沿与定时器每拍无条件刷新（禁置于 IF/CASE 内，使能挂 IN 引脚） —— *)
rtReset(CLK := bReset);
rtStart(CLK := bStart);
tonOpen (IN := (_ePhase = E_DL_SprayPhase.eOpen)  AND (NOT _bFault), PT := tOpen);
tonSpray(IN := (_ePhase = E_DL_SprayPhase.eSpray) AND (NOT _bFault), PT := tSpray);
tonBlow (IN := (_ePhase = E_DL_SprayPhase.eBlow)  AND (NOT _bFault), PT := tBlow);
tonClose(IN := (_ePhase = E_DL_SprayPhase.eClose) AND (NOT _bFault), PT := tClose);

(* —— 段 1｜每拍量预清零（锁存量 _bFault/_uFault/nSprayDone 不入清单） —— *)
uErrId := 16#0000_0000;
_bCfgBad := FALSE;

(* —— 段 2｜复位沿：故障一次性清干净，相位回空闲，喷涂计数清零 —— *)
IF rtReset.Q THEN
    _bFault := FALSE;
    _uFault := 16#0000_0000;
    nSprayDone := 0;
    _ePhase := E_DL_SprayPhase.eIdle;
END_IF

(* —— 段 3｜组态闸：喷涂次数与四段时长全覆盖 —— *)
IF (nSpraySet < 1) OR (tOpen = T#0S) OR (tSpray = T#0S) OR (tBlow = T#0S) OR (tClose = T#0S) THEN
    _bCfgBad := TRUE;
END_IF

(* —— 段 4｜主状态机：七态全覆盖 + ELSE 兜底 —— *)
CASE _ePhase OF
E_DL_SprayPhase.eIdle:
    bOpenCmd := FALSE; bSprayCmd := FALSE; bBlowCmd := FALSE; bCloseCmd := FALSE;
    IF rtStart.Q AND bEnable AND (NOT _bFault) AND (NOT _bCfgBad) THEN
        nSprayDone := 0;
        _ePhase := E_DL_SprayPhase.eOpen;
    ELSIF rtStart.Q AND (_bFault OR _bCfgBad) THEN
        _bFault := TRUE;                 (* 带病启动拒绝 / Reject start with bad config *)
        _uFault := 16#0025_0001;
        _ePhase := E_DL_SprayPhase.eFault;
    END_IF

E_DL_SprayPhase.eOpen:
    bOpenCmd := TRUE; bSprayCmd := FALSE; bBlowCmd := FALSE; bCloseCmd := FALSE;
    IF tonOpen.Q THEN
        _ePhase := E_DL_SprayPhase.eSpray;   (* 迁出条件 1：开模到位 *)
    ELSIF NOT bEnable THEN
        _ePhase := E_DL_SprayPhase.eIdle;    (* 迁出条件 2：使能撤销回安全态 *)
    END_IF

E_DL_SprayPhase.eSpray:
    bOpenCmd := TRUE; bSprayCmd := TRUE; bBlowCmd := FALSE; bCloseCmd := FALSE;
    IF tonSpray.Q THEN
        nSprayDone := nSprayDone + 1;        (* 次数在迁出拍单点累加 *)
        _ePhase := E_DL_SprayPhase.eBlow;    (* 迁出条件 1：单次喷涂完成 *)
    ELSIF NOT bEnable THEN
        _ePhase := E_DL_SprayPhase.eIdle;    (* 迁出条件 2：使能撤销 *)
    END_IF

E_DL_SprayPhase.eBlow:
    bOpenCmd := TRUE; bSprayCmd := FALSE; bBlowCmd := TRUE; bCloseCmd := FALSE;
    IF tonBlow.Q THEN
        IF nSprayDone < nSpraySet THEN
            _ePhase := E_DL_SprayPhase.eSpray;   (* 次数未达：重复喷涂-吹扫 *)
        ELSE
            _ePhase := E_DL_SprayPhase.eClose;   (* 迁出条件 1：次数达成转关模 *)
        END_IF
    ELSIF NOT bEnable THEN
        _ePhase := E_DL_SprayPhase.eIdle;        (* 迁出条件 2：使能撤销 *)
    END_IF

E_DL_SprayPhase.eClose:
    bOpenCmd := FALSE; bSprayCmd := FALSE; bBlowCmd := FALSE; bCloseCmd := TRUE;
    IF tonClose.Q THEN
        _ePhase := E_DL_SprayPhase.eDone;    (* 迁出条件 1：关模到位 *)
    ELSIF NOT bEnable THEN
        _ePhase := E_DL_SprayPhase.eIdle;    (* 迁出条件 2：使能撤销 *)
    END_IF

E_DL_SprayPhase.eDone:
    bOpenCmd := FALSE; bSprayCmd := FALSE; bBlowCmd := FALSE; bCloseCmd := FALSE;
    IF NOT bStart THEN
        _ePhase := E_DL_SprayPhase.eIdle;    (* 启动指令撤销：回空闲 *)
    END_IF

E_DL_SprayPhase.eFault:
    bOpenCmd := FALSE; bSprayCmd := FALSE; bBlowCmd := FALSE; bCloseCmd := FALSE;

ELSE
    _bFault := TRUE;                         (* 兜底：非法相位锁存 *)
    _uFault := 16#0025_0009;
    _ePhase := E_DL_SprayPhase.eFault;
END_CASE

(* —— 段 5｜相位与故障码出口单点映射 —— *)
ePhase := _ePhase;
bError := _bFault;
IF _bFault AND (_uFault <> 16#0000_0000) THEN
    uErrId := _uFault;                       (* 故障码锁存回放 / Latched fault replay *)
END_IF
END_FUNCTION_BLOCK

(* ---- FB_DL_DolMotor.st ---- *)
(*==============================================================================
 * 组件名称 (Component)  : FB_DL_DolMotor
 * 所属子库 (Sublibrary) : DL_Device
 * 当前版本 (Version)    : 1.0.0
 * 兼容性   (Platform)   : CODESYS 3.5 / TwinCAT 3 / 汇川 InoProShop / Machine Expert
 *                         仅依赖 Standard.library（TON / R_TRIG），零厂商方言
 * 分类     (Category)   : 设备执行器功能块（Function Block，实现 I_DL_MotorDriver）
 * 功能简述 (Function)   : 直接启动（DOL）电机控制功能块。含指令-反馈校验窗
 *                         （拒动保护）、运行失反馈脱扣、热继电器过载锁存、
 *                         最短运行时间监视、60 分钟桶滑窗每小时启动次数
 *                         限制与停机后重启抑制冷却；状态机采用
 *                         ENUM + CASE + ELSE 兜底。
 * 接口实现 (Implements) : I_DL_MotorDriver（属性 eState/bRunning/bFault/
 *                         uErrorId/bRestartInhibit，方法 CmdStart/CmdStop/
 *                         CmdReset，全部在本文件尾部落地）
 * 开源溯源 (Origin)     : 来源标签 lbp-device（RAW_NOTES_R5 S-4：DOL 电机侧
 *                         接触器反馈校验（指令-反馈 500ms 窗）、热继电器
 *                         过载锁存、防频繁启停（重启抑制冷却时间）等行业
 *                         公知语义，公开教学资料，仅借鉴通用工程语义；
 *                         状态机、小时窗计数算法、故障码按本库红线独立
 *                         设计，clean-room 未复制源码）。
 * 红线自检 (Redline)    : R1 零全局变量表/外部变量引用 ✓｜R2 零物理 IO 地址 ✓
 *                         R3 纯 IEC 61131-3 ✓｜R4 数组上下界防御+无死循环 ✓
 *                         R5 全变量中英双语同行注释 ✓｜R6 ENUM+CASE+ELSE ✓
 *                         R7 定时器/边缘实例主体最前部无条件刷新 ✓
 * 公约遵循 (Convention) : 0.1 本块为纯事件型状态机，无积分/滤波类首扫初始化
 *                         逻辑（分钟桶数组零值初始化由编译器缺省保证），
 *                         首扫跟踪范式不适用，无内部初始化标志。
 *                         0.7 故障码段位 16#0003_xxxx：【故障级】0003_0205
 *                         接触器拒动 / 0003_0206 失反馈脱扣 / 0003_0209
 *                         过载锁存 / 0003_0201 非法状态（全部 R15 锁存仅
 *                         复位可清）；【信息级】0003_0207 每小时启动次数
 *                         超限拒绝 / 0003_0208 重启抑制期拒绝 / 0003_020A
 *                         最短运行时间不足（仅写 uErrorId，不进 bFault，
 *                         0.2 公约）。
 * 修订历史 (Revision)   :
 *   2026-11-15  v1.0.0  首版入库（R5 轮 · DL_Device 开库）
 *============================================================================*)
FUNCTION_BLOCK FB_DL_DolMotor IMPLEMENTS I_DL_MotorDriver
VAR_INPUT
    bCmdStart         : BOOL;           // 启动指令（Start command），上升沿生效 / Start command, rising edge effective
    bCmdStop          : BOOL;           // 停止指令（Stop command），电平生效 / Stop command, level effective
    bFbContactor      : BOOL;           // 接触器辅助触点反馈（Contactor feedback），TRUE=吸合 / Contactor feedback, TRUE = picked up
    bThermalOverload  : BOOL;           // 热继电器过载信号（Thermal overload trip），TRUE=过载 / Thermal overload trip, TRUE = overloaded
    bPermitStart      : BOOL;           // 启动允许联锁（Start permit），TRUE=允许 / Start permit interlock, TRUE = start allowed
    tFbWindow         : TIME := T#500MS; // 指令-反馈校验窗口（Feedback check window），T#0S=免校验 / Feedback check window, T#0S disables the check
    tMinRunTime       : TIME := T#5S;   // 最短运行时间（Min run time），T#0S=免监视 / Minimum run time, T#0S disables the monitor
    tRestartInhibit   : TIME := T#60S;  // 重启抑制冷却时间（Restart inhibit），停机后冷却期内拒绝启动 / Restart inhibit cooling time after stop
    uMaxStartsPerHour : USINT := 6;     // 每小时最大启动次数（Max starts per hour），滑动小时窗上限 / Max starts per sliding hour window
    bReset            : BOOL;           // 故障复位（Fault reset），上升沿生效 / Fault reset, rising edge effective
END_VAR

VAR_OUTPUT
    bContactorCmd     : BOOL;           // 接触器线圈输出（Contactor coil command），TRUE=得电 / Contactor coil command, TRUE = energized
    eState            : E_DL_MotorState; // 当前状态机状态（Current state），映射接口同名属性 / Current state, mirrors interface property
    bRunning          : BOOL;           // 运行反馈（Running feedback），运行态且触点吸合确认 / Running feedback, running state confirmed by contactor
    bFault            : BOOL;           // 故障锁存中（Fault latched），TRUE=需复位 / Fault latched, TRUE requires reset
    uErrorId          : UDINT;          // 末次故障码（Last error code），0=无故障，段位 16#0003_xxxx / Last error code, 0 = none, family 16#0003_xxxx
    bRestartInhibit   : BOOL;           // 重启抑制激活中（Restart inhibit active），TRUE=冷却期拒绝启动 / Restart inhibit active, TRUE = starts refused
    uStartCount       : UDINT;          // 累计启动次数（Start count），每次受理启动 +1 / Total start count, incremented per accepted start
END_VAR

VAR
    _eState           : E_DL_MotorState := E_DL_MotorState.eIdle; // 内部状态机步序（Internal state step），外部经属性只读 / Internal state, read-only via property
    _bFaultLatch      : BOOL;           // 故障锁存标志（Fault latch flag），仅复位清除 / Fault latch flag, cleared only by reset
    _uErrorIdInt      : UDINT;          // 内部故障码寄存（Internal error register），故障级与信息级共用 / Internal error register, fault and info codes share it
    _bCooling         : BOOL;           // 冷却计时进行中（Cooling timing active）/ Cooling timer run request flag
    _bRestartInhibitAct : BOOL;         // 重启抑制激活内部寄存（Internal restart inhibit register）/ Internal restart inhibit register
    _bStopLatch       : BOOL;           // 方法停止锁存（Method stop latch），电平语义至回空闲态消化 / Method stop latch, level semantics until idle
    _bPendStart       : BOOL;           // 方法启动请求（Method start request），由 CmdStart 置位 / Method start request set by CmdStart
    _bPendReset       : BOOL;           // 方法复位请求（Method reset request），由 CmdReset 置位 / Method reset request set by CmdReset
    _bFbWinEn         : BOOL;           // 反馈校验窗使能（Feedback window enable），窗口参数大于零时有效 / Feedback window enable, active when window above zero
    _bMinRunEn        : BOOL;           // 最短运行监视使能（Min run monitor enable），参数大于零时有效 / Min run monitor enable, active when parameter above zero
    _bTickReset       : BOOL;           // 分钟桶定时器单周期复位保持（One-cycle tick timer hold-down）/ One-cycle hold-down to restart minute tick timer
    _aMinuteStarts    : ARRAY[0..59] OF UDINT; // 60 分钟启动次数桶（Sliding 60-minute start buckets），索引 0=当前分钟槽 / Buckets of starts per minute, index 0 = current slot
    _uMinIdx          : UINT;           // 当前分钟桶索引（Current minute bucket index），0..59 循环 / Current minute bucket index, cyclic 0..59
    _uHourCount       : UDINT;          // 滑动小时窗合计启动次数（Sliding hour window start sum）/ Start sum over sliding hour window
    _fbTrigStart      : R_TRIG;         // 引脚启动指令上升沿（Pin start command edge）/ Pin start command rising edge
    _fbTrigReset      : R_TRIG;         // 引脚复位上升沿（Pin reset edge）/ Pin reset rising edge
    _fbTrigTick       : R_TRIG;         // 分钟桶滚动触发（Minute bucket roll trigger）/ Minute bucket roll edge trigger
    _fbTonFbWindow    : TON;            // 指令-反馈校验窗定时器（Feedback check window timer）/ Feedback check window timer
    _fbTonMinRun      : TON;            // 最短运行时间定时器（Min run time timer）/ Minimum run time timer
    _fbTonRestartInh  : TON;            // 重启抑制冷却定时器（Restart inhibit cooling timer）/ Restart inhibit cooling timer
    _fbTonHourTick    : TON;            // 分钟桶节拍定时器（Minute tick timer），60 秒滚动 / Minute tick timer, rolls every 60 s
    i                 : UINT;           // 滑窗求和循环索引（Sliding window sum loop index）/ Loop index for window sum
END_VAR

METHOD CmdStart : BOOL
VAR_INPUT
END_VAR
IF (_eState <> E_DL_MotorState.eIdle) OR _bFaultLatch OR _bRestartInhibitAct THEN
    CmdStart := FALSE;        // 非空闲/故障/冷却期拒绝（Refused: not idle, faulty, or cooling）
ELSE
    _bPendStart := TRUE;      // 登记启动请求，主体状态机评估（Register start request, evaluated by body）
    CmdStart    := TRUE;      // 受理成功（Accepted）
END_IF

(*------------------------------------------------------------------------------
 * 方法: CmdStop —— 无条件安全停止（双线圈全断语义，由主体在运行/启动态消化）。
 *      Method CmdStop - unconditional safe stop, consumed by body in running/starting.
 *------------------------------------------------------------------------------*)
    END_METHOD

METHOD CmdStop
VAR_INPUT
END_VAR
_bStopLatch := TRUE;          // 登记停止锁存，主体状态机消化（Register stop latch, consumed by body）

(*------------------------------------------------------------------------------
 * 方法: CmdReset —— 复位过载/故障，返回是否可复位（存在锁存故障时为 TRUE）。
 *      Method CmdReset - reset overload/fault, returns TRUE only when latch exists.
 *------------------------------------------------------------------------------*)
    END_METHOD

METHOD CmdReset : BOOL
VAR_INPUT
END_VAR
IF _bFaultLatch OR (_eState = E_DL_MotorState.eFault) OR (_eState = E_DL_MotorState.eTripOverload) THEN
    _bPendReset := TRUE;      // 登记复位请求，主体状态机消化（Register reset request, consumed by body）
    CmdReset    := TRUE;      // 可复位（Resettable）
ELSE
    CmdReset    := FALSE;     // 无故障可复位（Nothing to reset）
END_IF

(*------------------------------------------------------------------------------
 * 属性: eState（GET）—— 当前状态机状态只读视图。
 *      Property eState (GET) - read-only view of the current state machine state.
 *------------------------------------------------------------------------------*)
    END_METHOD

// ============================================================================
// 段 1｜定时器与边缘检测实例无条件周期刷新（R7：严禁置于 IF/CASE 分支内）
//      Unconditional per-cycle refresh of all timer and edge instances (R7)
// ============================================================================
_fbTrigStart(CLK := bCmdStart);
_fbTrigReset(CLK := bReset);
_bFbWinEn := (tFbWindow > T#0S);    // 窗口为零 = 免校验（Zero window = check disabled）
_bMinRunEn := (tMinRunTime > T#0S); // 参数为零 = 免监视（Zero parameter = monitor disabled）
_fbTonFbWindow(IN := (_eState = E_DL_MotorState.eStarting) AND _bFbWinEn, PT := tFbWindow);
_fbTonMinRun(IN := ((_eState = E_DL_MotorState.eStarting) OR (_eState = E_DL_MotorState.eRunning)) AND _bMinRunEn, PT := tMinRunTime);
_fbTonRestartInh(IN := _bCooling, PT := tRestartInhibit);
_fbTonHourTick(IN := NOT _bTickReset, PT := T#60S);
_fbTrigTick(CLK := _fbTonHourTick.Q);

// 冷却到期：解除抑制（Cooling expired: release inhibit）
IF _fbTonRestartInh.Q THEN
    _bCooling           := FALSE;    // 结束冷却计时（Stop cooling timing）
    _bRestartInhibitAct := FALSE;    // 解除抑制（Release inhibit）
ELSE
    _bRestartInhibitAct := _bCooling; // 冷却期间抑制有效（Inhibit active during cooling）
END_IF

// ============================================================================
// 段 2｜滑动小时窗：60 秒滚动分钟桶 + 全窗求和（固定界 FOR，无死循环风险）
//      Sliding hour window: 60 s rolling minute buckets + full window sum
// ============================================================================
IF _fbTrigTick.Q THEN
    _uMinIdx := (_uMinIdx + 1) MOD 60; // 桶索引循环推进（Advance bucket index cyclically）
    IF _uMinIdx <= 59 THEN
        _aMinuteStarts[_uMinIdx] := 0; // 新槽清零，旧数据保留 59 分钟后自然滑出（Clear new slot, old data slides out after 59 min）
    END_IF
    _bTickReset := TRUE;               // 单周期复位节拍定时器（One-cycle reset of tick timer）
END_IF
IF _bTickReset THEN
    _bTickReset := FALSE;              // 下一周期恢复计时（Resume timing next cycle）
END_IF

_uHourCount := 0;                      // 每周期重算滑窗合计（Recompute window sum each cycle）
FOR i := 0 TO 59 DO
    _uHourCount := _uHourCount + _aMinuteStarts[i]; // 累加 60 个分钟桶（Accumulate all 60 buckets）
END_FOR

// ============================================================================
// 段 3｜过载全局监视（优先级最高）：启动/运行态过载立即锁存脱扣
//      Global overload monitor (highest priority): trip immediately in starting/running
// ============================================================================
IF bThermalOverload AND ((_eState = E_DL_MotorState.eStarting) OR (_eState = E_DL_MotorState.eRunning)) THEN
    _bFaultLatch := TRUE;              // 过载锁存（Overload latched）
    _uErrorIdInt := 16#0003_0209;      // 0003_0209 热继电器过载脱扣【故障级】/ Thermal overload trip, fault level
    _eState      := E_DL_MotorState.eTripOverload; // 强制脱扣态（Force trip state）
END_IF

// ============================================================================
// 段 4｜核心状态机（ENUM + CASE，含 ELSE 非法状态兜底）
//      Core state machine (ENUM + CASE with ELSE illegal-state fallback)
// ============================================================================
CASE _eState OF

    E_DL_MotorState.eIdle: // 空闲停机态：消化停止锁存，评估启动请求
        IF _bStopLatch THEN
            _bStopLatch := FALSE;      // 停止锁存到空闲即消化（Stop latch absorbed at idle）
        END_IF
        IF _bPendStart OR _fbTrigStart.Q THEN
            IF bThermalOverload THEN
                _bPendStart := FALSE;  // 过载未复位：静默拒绝（Overload present: silent refusal, trip code already latched in trip state）
            ELSIF NOT bPermitStart THEN
                _bPendStart := FALSE;  // 联锁未满足：静默拒绝（Permit absent: silent refusal）
            ELSIF _bRestartInhibitAct THEN
                _bPendStart := FALSE;  // 消费请求不自动重试（Consume request, no auto retry）
                _uErrorIdInt := 16#0003_0208; // 0003_0208 重启抑制期内启动被拒【信息级】/ Start refused during restart inhibit, info level
            ELSIF _uHourCount >= uMaxStartsPerHour THEN
                _bPendStart := FALSE;  // 消费请求不自动重试（Consume request, no auto retry）
                _uErrorIdInt := 16#0003_0207; // 0003_0207 每小时启动次数超限拒绝【信息级】/ Hourly start limit exceeded, info level
            ELSE
                _bPendStart := FALSE;  // 受理启动（Accept start）
                uStartCount := uStartCount + 1; // 累计启动 +1（Total starts +1）
                IF _uMinIdx <= 59 THEN
                    _aMinuteStarts[_uMinIdx] := _aMinuteStarts[_uMinIdx] + 1; // 当前分钟桶 +1（Current bucket +1）
                END_IF
                _eState := E_DL_MotorState.eStarting;
            END_IF
        END_IF

    E_DL_MotorState.eStarting: // 启动校验态：线圈得电，等待反馈窗内吸合
        IF bFbContactor THEN
            _eState := E_DL_MotorState.eRunning;   // 吸合确认，转运行（Pick-up confirmed, to running）
        ELSIF _fbTonFbWindow.Q THEN
            _bFaultLatch := TRUE;                  // 拒动故障锁存（Refusal fault latch）
            _uErrorIdInt := 16#0003_0205;          // 0003_0205 接触器拒动（窗内未吸合）【故障级】/ Contactor refused to pick up in window, fault level
            _eState      := E_DL_MotorState.eFault;
        ELSIF bCmdStop OR _bStopLatch THEN
            _eState := E_DL_MotorState.eStopping;  // 启动中止：线圈断开，无运行故不计 0003_020A / Aborted start: no run time, 0003_020A not applicable
        END_IF

    E_DL_MotorState.eRunning: // 运行态：反馈吸合确认
        IF bCmdStop OR _bStopLatch THEN
            IF (NOT _fbTonMinRun.Q) AND _bMinRunEn THEN
                _uErrorIdInt := 16#0003_020A;      // 0003_020A 运行不足最短时间即停【信息级】/ Stopped before min run time, info level
            END_IF
            _eState := E_DL_MotorState.eStopping;  // 转停机过渡（To stopping transition）
        ELSIF NOT bFbContactor THEN
            _bFaultLatch := TRUE;                  // 失反馈脱扣锁存（Feedback loss latch）
            _uErrorIdInt := 16#0003_0206;          // 0003_0206 运行中反馈意外断开【故障级】/ Contactor feedback dropped while running, fault level
            _eState      := E_DL_MotorState.eFault;
        END_IF

    E_DL_MotorState.eStopping: // 停机过渡态：线圈已断，等反馈分断
        IF NOT bFbContactor THEN
            _bStopLatch := FALSE;                  // 停止锁存消化（Stop latch absorbed）
            _bCooling   := TRUE;                   // 启动重启抑制冷却（Start restart-inhibit cooling）
            _eState     := E_DL_MotorState.eIdle;  // 回空闲（Back to idle）
        END_IF
        // 反馈触点粘连时保持本态等待分断，直至上层干预（Welded contact holds this state until intervention）

    E_DL_MotorState.eTripOverload: // 过载脱扣锁存态：仅复位且过载消失后可清
        IF (_fbTrigReset.Q OR _bPendReset) AND (NOT bThermalOverload) THEN
            _bPendReset  := FALSE;                 // 消费复位请求（Consume reset request）
            _bFaultLatch := FALSE;                 // 解除锁存（Release latch）
            _uErrorIdInt := 0;                     // 故障码清零（Error code cleared）
            _bCooling    := TRUE;                  // 脱扣复位后同样进入冷却（Cooling also after trip reset）
            _eState      := E_DL_MotorState.eIdle; // 回空闲（Back to idle）
        END_IF

    E_DL_MotorState.eFault: // 故障锁存态：仅复位可退出
        IF _fbTrigReset.Q OR _bPendReset THEN
            _bPendReset  := FALSE;                 // 消费复位请求（Consume reset request）
            _bFaultLatch := FALSE;                 // 解除锁存（Release latch）
            _uErrorIdInt := 0;                     // 故障码清零（Error code cleared）
            _bCooling    := TRUE;                  // 故障复位后进入冷却（Cooling also after fault reset）
            _eState      := E_DL_MotorState.eIdle; // 回空闲（Back to idle）
        END_IF

    ELSE // 非法状态兜底：任何越界枚举值强制锁存故障（Illegal state fallback）
        _bFaultLatch := TRUE;                      // 故障锁存（Fault latched）
        _uErrorIdInt := 16#0003_0201;              // 0003_0201 非法状态【故障级】/ Illegal state, fault level
        _eState      := E_DL_MotorState.eFault;
END_CASE

// ============================================================================
// 段 5｜输出映射（bFault 为显式派生式：仅故障级码可达的锁存/状态置位，
//         信息级 0003_0207/0208/020A 天然被排除——0.2 公约）
//      Output mapping (bFault explicit derived form: only fault-level codes
//      can set it, info codes 0003_0207/0208/020A excluded by construction)
// ============================================================================
bContactorCmd   := (_eState = E_DL_MotorState.eStarting) OR (_eState = E_DL_MotorState.eRunning); // 仅启动/运行态得电（Energized only in starting/running）
eState          := _eState;                       // 状态映射（State mapping）
bRunning        := (_eState = E_DL_MotorState.eRunning) AND bFbContactor; // 运行 = 状态且反馈确认（Running = state AND feedback confirmed）
bFault          := _bFaultLatch OR (_eState = E_DL_MotorState.eFault) OR (_eState = E_DL_MotorState.eTripOverload); // 故障派生（Fault derived）
uErrorId        := _uErrorIdInt;                  // 故障码映射（Error code mapping）
bRestartInhibit := _bRestartInhibitAct;           // 重启抑制映射（Restart inhibit mapping）

(*------------------------------------------------------------------------------
 * 方法: CmdStart —— 启动指令（单发）。被抑制（冷却中）或故障态返回 FALSE。
 *      Method CmdStart - start command (one-shot), FALSE when inhibited or faulty.
 *------------------------------------------------------------------------------*)

PROPERTY eState : E_DL_MotorState
eState := _eState;            // 返回内部状态（Return internal state）

(*------------------------------------------------------------------------------
 * 属性: bRunning（GET）—— 运行反馈（状态且触点吸合确认）。
 *      Property bRunning (GET) - running feedback (state AND contactor confirmed).
 *------------------------------------------------------------------------------*)
PROPERTY bRunning : BOOL
bRunning := (_eState = E_DL_MotorState.eRunning) AND bFbContactor; // 显式确认式派生（Explicit confirmed derived form）

(*------------------------------------------------------------------------------
 * 属性: bFault（GET）—— 故障锁存指示（信息级码不置本位，0.2 公约）。
 *      Property bFault (GET) - fault latch indicator, info-level codes excluded.
 *------------------------------------------------------------------------------*)
PROPERTY bFault : BOOL
bFault := _bFaultLatch OR (_eState = E_DL_MotorState.eFault) OR (_eState = E_DL_MotorState.eTripOverload); // 显式排除信息级派生式（Explicit derived form excluding info codes）

(*------------------------------------------------------------------------------
 * 属性: uErrorId（GET）—— 末次故障码（0=无故障）。
 *      Property uErrorId (GET) - last error code (0 = none).
 *------------------------------------------------------------------------------*)
PROPERTY uErrorId : UDINT
uErrorId := _uErrorIdInt;     // 返回内部故障码寄存（Return internal error register）

(*------------------------------------------------------------------------------
 * 属性: bRestartInhibit（GET）—— 重启抑制激活指示。
 *      Property bRestartInhibit (GET) - restart inhibit active indicator.
 *------------------------------------------------------------------------------*)
PROPERTY bRestartInhibit : BOOL
bRestartInhibit := _bRestartInhibitAct; // 返回抑制寄存（Return inhibit register）
END_FUNCTION_BLOCK

(* ---- FB_DL_DoorInterlockHvac.st ---- *)
(*
  FB_DL_DoorInterlockHvac  —  机房门禁-风机联锁（开门降频 → 关门延时恢复）/ Door interlock with fan speed ramp-down
  分类 Category : DL_Device
  码位 Code     : 16#03_2_18
  段位说明      : 03_2 段低半字节已满，1x 段续号，17 格由 BcdFieldPanelIO 启用，本件启用 18 格（R192）
  版本 Version  : 1.0.0
  来源 Source   : t2-2-lbp — 门禁-风机「降频-恢复」策略组态待挖项
  溯源 Origin   : clean-room 实现，未复制任何源码行
                  （与 FB_DL_GuardLockDoor 分工：那件管门本体握手；与炉门互锁族分工：那族管全停互锁，
                   本件管「降频-恢复」而非全停——风机保持运行仅限速，保障机房排风）
  功能 Function : 1) 四相联锁 Normal→Reduced→RestoreWait→Normal：开门（消抖/模拟量迟滞双口径）
                  降频至 fDoorOpenSpdPct，关门后经 tRestoreDelay 延时恢复需求转速；
                  2) 降频目标经 FB_DL_RateLimiter 斜坡（fRateUpPctS/fRateDownPctS 分向速率），
                  风机不失电不喘振；
                  3) 模拟量门磁口径（bUseAnaDoor = TRUE）：门缝宽度经 FC_DL_Hysteresis 迟滞判门态；
                  数字量口径：经 FB_DL_SignalDebounce 消抖判门态；
                  4) 故障相（组态非法）风机指令强制归零（安全侧：机房排风联锁失效宁可停风机报警）。
  边界 Boundary : ① 本件只出转速指令 fFanSpdCmdPct，不写风机本体 IO（由上层 PRG_IoMapping 承载）；
                  ② 门开降频与关门恢复的策略参数（速率/延时/降频值）全部引脚化组态；
                  ③ R228-A 达标声明：tonRestore 单相独占（IN 为单相等式），跨相迁移拍 IN 必断；
                  ④ R228-B 达标声明：eFault 迁出 = rtReset.Q（输入引脚，恒可达），逐字写于此；
                  ⑤ 迟滞判门态时 fDoorHystMm 越组态域按上限钳位（防御误填，不中断扫描）。
  依赖 Depends  : FB_DL_RateLimiter / FB_DL_SignalDebounce（实例化，引脚按 registry 实名）；
                  FC_DL_Hysteresis（函数调用，bState 由本件成员持有回传）
  码表 Error codes（本件格 03_2_18，子码步进 +0x100）:
    16#0003_0118 信息级：降频目标已到达（Reduced 相稳定）
    16#0003_0218 故障级：组态非法（需求/降频值越 0..100 / 速率非法 / 迟滞域非法），锁存至复位
    16#0003_0318 信息级：关门恢复延时进行中（RestoreWait 相，不置故障）
    16#0003_0418 故障级：状态机落 ELSE 兜底（非法相位 ID），锁存至复位

  修订历史 Revision :
    2026-11-19  v1.0.0  R39 首版（批次 2 · 序号 10）
*)

TYPE E_DL_DoorIntState :
(
    eNormal      := 0,    // 正常：需求转速直通 / Normal, demand speed passes through
    eReduced     := 10,   // 降频：门开，指令钳到降频值 / Reduced, door open, speed clamped
    eRestoreWait := 20,   // 恢复等待：门关，延时恢复 / Restore wait, door closed, delayed restore
    eFault       := 90    // 故障：组态锁定，指令归零 / Fault, latched, command forced to zero
);
END_TYPE

FUNCTION_BLOCK FB_DL_DoorInterlockHvac
VAR_INPUT
    bEnable         : BOOL := TRUE;       // 总使能，FALSE 时指令归零并回 Normal 判定冻结 [-] / Master enable
    bDoorOpenRaw    : BOOL := FALSE;      // 数字量门磁原始信号（bUseAnaDoor = FALSE 时生效）/ Digital door switch raw input
    fDoorGapMm      : REAL := 0.0;        // 模拟量门缝宽度 [mm]（bUseAnaDoor = TRUE 时生效）/ Analog door gap width
    bUseAnaDoor     : BOOL := FALSE;      // 门态判据口径选择：TRUE = 模拟量迟滞 / FALSE = 数字消抖 / Door sensing mode select
    fDoorThrMm      : REAL := 30.0;       // 门缝开门判据阈 [mm]，域 > 0 / Analog door-open threshold
    fDoorHystMm     : REAL := 5.0;        // 门缝迟滞带 [mm]，域 > 0 / Analog door hysteresis band
    fFanSpdReqPct   : REAL := 80.0;       // 正常需求转速 [%]，域 [0, 100] / Normal demand speed
    fDoorOpenSpdPct : REAL := 30.0;       // 门开降频转速 [%]，域 [0, 100] / Door-open reduced speed
    fRateUpPctS     : REAL := 20.0;       // 恢复上升速率 [%/s]，域 > 0 / Restore ramp-up rate
    fRateDownPctS   : REAL := 40.0;       // 降频下降速率 [%/s]，域 > 0 / Reduced ramp-down rate
    tRestoreDelay   : TIME := T#5S;       // 关门恢复延时 [ms]，域 > 0 / Restore delay after door closed
    tSampleTime     : TIME := T#100MS;    // 限速器采样周期 [ms] / Rate limiter sample period
    bReset          : BOOL := FALSE;      // 故障复位，上升沿生效 / Fault reset, rising edge
END_VAR
VAR_OUTPUT
    fFanSpdCmdPct : REAL;                 // 风机转速指令 [%]（上层风机消费）/ Fan speed command output
    bDoorDeb      : BOOL;                 // 门态判定出口（消抖/迟滞后）/ Judged door state output
    bReduced      : BOOL;                 // 降频生效中（Reduced 相）[-] / Reduced mode active
    bRestorePend  : BOOL;                 // 恢复延时进行中（RestoreWait 相）[-] / Restore delay in progress
    eState        : E_DL_DoorIntState;    // 状态出口，段尾单点映射 / State outlet
    bError        : BOOL;                 // 故障锁存，仅故障级码置位，bReset 清除 [-] / Fault latch
    uErrorId      : UDINT;                // 事件码，0 = 无事件（故障级锁存回放）/ Event code
END_VAR
VAR
    fbDeb       : FB_DL_SignalDebounce;   // 数字量门磁消抖实例（主体首部无条件刷新）/ Digital door debounce instance
    fbLim       : FB_DL_RateLimiter;      // 转速斜坡限速实例（主体首部无条件刷新）/ Speed ramp limiter instance
    tonRestore  : TON;                    // 恢复延时计时（单相独占，R228-A）/ Restore delay timer, single phase
    rtReset     : R_TRIG;                 // 复位上升沿 / Reset rising edge
    _eState     : E_DL_DoorIntState := E_DL_DoorIntState.eNormal;  // 内部相位（CASE 唯一写入目标）/ Internal phase
    _bDoorSt    : BOOL;                   // 迟滞判门态回传保持变量（FC_DL_Hysteresis 有状态纪律）/ Hysteresis door-state hold member
    _rTarget    : REAL;                   // 本拍目标转速 [%] / Target speed this cycle
    _rDoorSpdEff: REAL := 30.0;           // 钳位后降频转速 [%] / Clamped reduced speed
    _rReqEff    : REAL := 80.0;           // 钳位后需求转速 [%] / Clamped demand speed
    _bFault     : BOOL;                   // 故障锁存位 / Latched fault bit
    _uFault     : UDINT;                  // 故障码锁存寄存 / Latched fault code register
    _uInfo      : UDINT;                  // 信息码，每拍重算 / Info code
    _bCfgBad    : BOOL;                   // 组态非法聚合 / Configuration invalid aggregate
END_VAR
VAR CONSTANT
    DL_DIH_INF_CAP : REAL := 1.0E15;    // 非有限值筛查幅值上限 / Non-finite screening cap
    DL_DIH_DT_MIN  : TIME := T#10MS;    // 限速器采样周期下限 [ms] / Rate limiter sample lower clamp
END_VAR

(* —— 段 0：定时器与边沿实例无条件周期刷新（R182：调用语句不得置于 IF/CASE 内） —— *)
rtReset(CLK := bReset);                                                 // 复位沿刷新，每拍必调
fbDeb(bRawInput := bDoorOpenRaw,                                        // 数字门磁消抖
      tRiseDelay := T#100MS,                                            // 上升确认延时（门磁标准口径）
      tFallDelay := T#100MS,                                            // 下降确认延时
      bEnable := NOT bUseAnaDoor);                                      // 数字口径使能（模拟口径旁路）
fbLim(bEnable := TRUE,                                                  // 限速器恒使能（跨相平滑）
      fIn := _rTarget,                                                  // 限速输入 = 本拍目标
      fRateUp := MAX(fRateUpPctS, 1.0E-6),                              // 上升速率（下限防零速率卡死）
      fRateDown := MAX(fRateDownPctS, 1.0E-6),                          // 下降速率（下限防零速率卡死）
      bTrack := FALSE,                                                  // 不跟踪（转速指令连续性优先）
      fTrackValue := 0.0,                                               // 跟踪值（未用，占位保持接口完整）
      tSampleTime := MAX(tSampleTime, DL_DIH_DT_MIN));                  // 采样周期（下限钳位）
tonRestore(IN := (_eState = E_DL_DoorIntState.eRestoreWait) AND (NOT bDoorSt), PT := tRestoreDelay);   // 恢复延时（单相独占）

(* —— 段 1：单拍量预清零（锁存量 _uFault/_bFault/_bDoorSt 不入清单，R187①） —— *)
_uInfo := 16#0000_0000;             // 信息码每拍重算
_bCfgBad := FALSE;                  // 组态非法预清零
_rTarget := 0.0;                    // 目标转速预清零（段 4 单点重写）

(* —— 段 2：组态域闸（覆盖全部参与判据换算的引脚，R151） —— *)
IF (fFanSpdReqPct < 0.0) OR (fFanSpdReqPct > 100.0)
   OR (fDoorOpenSpdPct < 0.0) OR (fDoorOpenSpdPct > 100.0)
   OR (fRateUpPctS <= 0.0) OR (fRateDownPctS <= 0.0)
   OR (TIME_TO_DINT(tRestoreDelay) <= 0) THEN
    _bCfgBad := TRUE;               // 需求/降频值越域或速率/延时非法
END_IF
IF (fDoorGapMm <> fDoorGapMm) OR (ABS(fDoorGapMm) > DL_DIH_INF_CAP) OR ((fDoorGapMm - fDoorGapMm) <> 0.0) THEN
    _bCfgBad := TRUE;               // 门缝输入非有限
END_IF
IF bUseAnaDoor AND ((fDoorThrMm <= 0.0) OR (fDoorHystMm <= 0.0) OR (fDoorHystMm > fDoorThrMm * 0.5)) THEN
    _bCfgBad := TRUE;               // 模拟口径阈值/迟滞非法（迟滞不越过阈值一半）
END_IF

(* —— 段 3：故障锁存与 eFault 迁出沿（R228-B：迁出条件 rtReset.Q 恒可达） —— *)
IF _bCfgBad AND (NOT _bFault) THEN
    _uFault := 16#0003_0218;        // 故障级：组态非法（仅首次进入时写入）
    _bFault := TRUE;
END_IF
IF rtReset.Q AND (NOT _bCfgBad) THEN
    _bFault := FALSE;               // 清故障锁存位（组态恢复合法为前提）
    _uFault := 16#0000_0000;
    IF _eState = E_DL_DoorIntState.eFault THEN
        _eState := E_DL_DoorIntState.eNormal;   // 故障相迁出：回正常相
    END_IF
END_IF

(* —— 段 4：门态判定与目标转速计算（故障相强制归零，安全侧） —— *)
_rReqEff := fFanSpdReqPct;          // 需求转速生效值（域已由段 2 闸门保证 0..100）
_rDoorSpdEff := fDoorOpenSpdPct;    // 降频转速生效值（域已由段 2 闸门保证 0..100）
IF bUseAnaDoor THEN
    bDoorDeb := FC_DL_Hysteresis(fIn := fDoorGapMm,             // 模拟口径：门缝迟滞判门态
                                 fThreshold := fDoorThrMm,      // 开门阈
                                 fHysteresis := fDoorHystMm,    // 迟滞带
                                 bState := _bDoorSt);           // 回传保持变量（同一成员，有状态纪律）
ELSE
    bDoorDeb := fbDeb.bStable;      // 数字口径：消抖稳定值
END_IF
IF _bFault OR (NOT bEnable) THEN
    _rTarget := 0.0;                // 故障/失能：指令目标归零（安全侧）
ELSIF bDoorDeb THEN
    _rTarget := MIN(_rReqEff, _rDoorSpdEff);    // 门开：需求与降频值取小（降频不高于需求）
ELSE
    _rTarget := _rReqEff;           // 门关：需求直通
END_IF

(* —— 段 5：相位机（只做相迁移与信息码；出口在段 7） —— *)
CASE _eState OF

E_DL_DoorIntState.eNormal:
    IF bDoorDeb THEN
        _eState := E_DL_DoorIntState.eReduced;      // 门开：进降频相
    END_IF

E_DL_DoorIntState.eReduced:
    IF bDoorDeb AND (_rTarget <= _rDoorSpdEff) THEN
        _uInfo := 16#0003_0118;     // 信息级：降频目标已到达（斜坡收敛）
    END_IF
    IF NOT bDoorDeb THEN
        _eState := E_DL_DoorIntState.eRestoreWait;  // 门关：进恢复等待相
    END_IF

E_DL_DoorIntState.eRestoreWait:
    bRestorePend := TRUE;           // 恢复延时进行中（相内重申）
    IF bDoorDeb THEN
        _eState := E_DL_DoorIntState.eReduced;      // 门复开：回降频相（延时计时随相断，R228-A）
    ELSIF tonRestore.Q THEN
        _eState := E_DL_DoorIntState.eNormal;       // 延时到点：回正常相
    END_IF

E_DL_DoorIntState.eFault:
    ;                               // 故障相：等复位沿（段 3 承载迁出）

ELSE
    _uFault := 16#0003_0418;        // 故障级：非法相位 ID 兜底
    _bFault := TRUE;
    _eState := E_DL_DoorIntState.eFault;    // 强制回故障相

END_CASE

(* —— 段 6：出口单点映射（名实同源；锁存码回放，禁同拍抹除） —— *)
fFanSpdCmdPct := fbLim.fOut;        // 转速指令 = 限速器输出（斜坡平滑口径）
bReduced := (_eState = E_DL_DoorIntState.eReduced);         // 降频生效中
bRestorePend := (_eState = E_DL_DoorIntState.eRestoreWait); // 恢复延时进行中（相外重写覆盖相内置位，口径统一）
IF _bFault THEN
    uErrorId := _uFault;            // 故障锁存码回放
    bError := TRUE;
ELSE
    uErrorId := _uInfo;             // 信息码
    bError := FALSE;
END_IF
eState := _eState;                  // 状态出口单点映射

END_FUNCTION_BLOCK

(* ---- FB_DL_DosingPumpCalib.st ---- *)
(*==============================================================================
 * 组件名称 (Component)  : FB_DL_DosingPumpCalib
 * 所属子库 (Sublibrary) : DL_Device
 * 前缀     (Prefix)     : FB_DL_
 * 当前版本 (Version)    : 1.0.0
 * 兼容性   (Platform)   : CODESYS 3.5 / TwinCAT 3 / 汇川 InoProShop / Schneider
 *                         Machine Expert；纯 IEC 61131-3（第 3 版），
 *                         仅依赖标准库 R_TRIG / ABS，零厂商方言
 * 作者     (Author)     : 道莅代码库 · PLC编程专家（R31）
 * 开源溯源 (Origin)     : 计量泵脉冲当量标定公开工艺语义（半导体/化工通用），
 *                         道莅 clean-room 防御性实现，未复制任何外部源码行
 * 功能描述 (Function)   : 计量泵标定与脉冲当量校验件。由标定容积与实测容积
 *                         反算实测当量（毫升每脉冲），与组态当量比偏差，
 *                         超差给出告警码并输出按偏差反向修正、夹在组态
 *                         0.5~2.0 倍带内的修正当量，供泵组态直接替换。
 * 状态机   (States)     : eIdle 待机 / eRun 单拍计算 / eDone 单拍完成脉冲 /
 *                         eFault 故障锁定（CASE 带 ELSE 兜底）。
 * 码位     (Codes)      : 16#0003_00F7 信息级：中止请求提示（不置 bError）
 *                         16#0003_00F8 故障级：样本不足（脉冲数低于下限）
 *                         16#0003_00F9 故障级：容积非法（标定/实测容积非有限
 *                                      或不大于零）
 *                         16#0003_00FA 故障级：组态当量非法（非有限或不大于零）
 *                         16#0003_00FB 告警级：当量偏差超差（仅告警不置
 *                                      bError，规格 §5.2 条目 6 优先于槽位
 *                                      通则，头注释留档）
 * 边界防错 (Boundary)   : 1 脉冲数低于下限判样本不足拒绝出结果；
 *                         2 组态当量非法或非有限锁故障并冻结输出（保持末次
 *                           有效值，禁零值覆盖）；
 *                         3 分母（脉冲数）为零防护：与样本不足同槽拒绝；
 *                         4 bAbort 立即清忙、不产出半结果、不置完成；
 *                         5 bDone 为新沿后单拍脉冲（R27 输出保持语义：
 *                           跨拍须清零）；
 *                         6 故障锁存的可达解除路径：下一次 bStart 上升沿
 *                           重新受理（故障态下仍受理启动，复位即重试）。
 * 修订历史 (Revision)   : 2026-11-18 v1.0.0 首版入库（R31 · 阶段三 · 序 7，
 *                         替代原 EscChuckCurrentMon 派单，见派单勘误 §5.2）
 *==============================================================================*)

(*------------------------------------------------------------------------------
 * 枚举: E_DL_DpcState（归属本功能块，同文件发布，全库唯一属主）
 *----------------------------------------------------------------------------*)
TYPE E_DL_DpcState :
(
    eIdle  := 0,    // 待机：等待启动沿 / Idle, waiting for start edge
    eRun   := 10,   // 计算态：单拍完成标定计算 / Run, calibration computed in one scan
    eDone  := 20,   // 完成态：单拍完成脉冲后回待机 / Done, one-scan pulse then idle
    eFault := 99    // 故障态：锁存等待重试 / Fault, latched awaiting retry
);
END_TYPE

(*==============================================================================
 * 功能块: FB_DL_DosingPumpCalib
 * 调用约定: 每个扫描周期无条件调用一次；标定数据经引脚单次注入。
 *==============================================================================*)
FUNCTION_BLOCK FB_DL_DosingPumpCalib
VAR_INPUT
    bStart             : BOOL := FALSE;  // 启动沿（含故障态重试受理）/ Start edge, also retries from fault
    bAbort             : BOOL := FALSE;  // 中止请求，任意拍生效 / Abort request, effective on any scan
    fCalVolumeMl       : REAL := 100.0;  // 标定容积 [毫升] / Calibration volume [mL]
    fMeasuredMl        : REAL := 0.0;    // 实测收集容积 [毫升] / Measured collected volume [mL]
    uPulseCount        : UDINT := 0;     // 标定脉冲总数 [个] / Total pulse count [count]
    fNominalMlPerPulse : REAL := 0.1;    // 组态当量 [毫升每脉冲] / Configured equivalent [mL per pulse]
    fTolPct            : REAL := 2.0;    // 偏差告警限 [百分数] / Deviation alarm limit [%]
    uMinPulses         : UDINT := 100;   // 最小样本脉冲数 [个] / Minimum sample pulse count [count]
END_VAR
VAR_OUTPUT
    bBusy              : BOOL;           // 忙标志（计算当拍）/ Busy flag during compute scan
    bDone              : BOOL;           // 完成单拍脉冲（R27）/ Done one-scan pulse
    bError             : BOOL;           // 故障标志，与故障级码配对（R45）/ Fault flag paired with fault codes
    fMeasuredMlPerPulse : REAL;          // 实测当量 [毫升每脉冲] / Measured equivalent [mL per pulse]
    fDeviationPct      : REAL;           // 当量偏差 [百分数] / Equivalent deviation [%]
    fCorrectedMlPerPulse : REAL;         // 修正当量（反向修正并夹带）[毫升每脉冲] / Corrected equivalent [mL per pulse]
    uErrorId           : UDINT;          // 错误码，0 = 无错 / Error code, 0 = none
END_VAR
VAR
    rTrigStart         : R_TRIG;         // 启动沿检测，每拍无条件刷新 / Start edge detector, refreshed every scan
    eState             : E_DL_DpcState;  // 内部状态机 / Internal state machine
    bVolOk             : BOOL;           // 容积对有效性 / Volume pair validity
    bNomOk             : BOOL;           // 组态当量有效性 / Nominal equivalent validity
    bCntOk             : BOOL;           // 样本量有效性 / Sample count validity
    fMeasEquiv         : REAL;           // 计算暂存实测当量 [毫升每脉冲] / Staged measured equivalent [mL per pulse]
    fDevPct            : REAL;           // 计算暂存偏差 [百分数] / Staged deviation [%]
    fCorrEquiv         : REAL;           // 计算暂存修正当量 [毫升每脉冲] / Staged corrected equivalent [mL per pulse]
    fNomAbs            : REAL;           // 组态当量幅值夹带基准 [毫升每脉冲] / Nominal magnitude clamp base [mL per pulse]
    uCodeLatch         : UDINT;          // 故障级锁存码 / Latched fault code
END_VAR
VAR CONSTANT
    DL_DPC_FIN  : REAL  := 1.0E30;       // REAL 有限幅值判界 / REAL finiteness magnitude bound
    DL_DPC_LO   : REAL  := 0.5;          // 修正当量夹带下限系数（组态倍数）/ Corrected clamp low factor
    DL_DPC_HI   : REAL  := 2.0;          // 修正当量夹带上限系数（组态倍数）/ Corrected clamp high factor
    DL_DPC_PCT  : REAL  := 100.0;        // 百分数换算系数 / Percent conversion factor
END_VAR

// ---- 段 1｜边沿实例无条件刷新（红线：禁入条件分支）----------------------------
rTrigStart(CLK := bStart);                            // 启动沿检测 / Start edge detection

// ---- 段 2｜中止请求：立即清忙、不产出半结果、不置完成（信息级提示）--------------
IF bAbort AND ((eState = eRun) OR (eState = eDone)) THEN
    eState    := eIdle;                               // 中止回待机 / Abort returns to idle
    bBusy     := FALSE;                               // 立即清忙 / Clear busy at once
    bDone     := FALSE;                               // 不置完成 / Never set done
    uErrorId  := 16#0003_00F7;                        // 信息级：中止提示 / Info: abort notice
END_IF

// ---- 段 3｜完成脉冲收尾（单拍语义，跨拍清零）------------------------------------
IF eState = eDone THEN
    bDone  := TRUE;                                   // 完成单拍脉冲 / One-scan done pulse
    bBusy  := FALSE;                                  // 完成态清忙 / Clear busy in done
    eState := eIdle;                                  // 下拍回待机 / Back to idle next scan
ELSIF eState = eRun THEN
    bBusy := TRUE;                                    // 计算当拍置忙 / Busy during compute scan
END_IF

// ---- 段 4｜启动沿受理（含故障态重试）--------------------------------------------
IF rTrigStart.Q AND ((eState = eIdle) OR (eState = eFault)) THEN
    bVolOk := (fCalVolumeMl = fCalVolumeMl) AND (fMeasuredMl = fMeasuredMl)
          AND (ABS(fCalVolumeMl) < DL_DPC_FIN) AND (ABS(fMeasuredMl) < DL_DPC_FIN)
          AND (fCalVolumeMl > 0.0) AND (fMeasuredMl > 0.0); // 容积对有限且大于零 / Volumes finite and positive
    bNomOk := (fNominalMlPerPulse = fNominalMlPerPulse)
          AND (ABS(fNominalMlPerPulse) < DL_DPC_FIN)
          AND (fNominalMlPerPulse > 0.0);             // 组态当量有限且大于零 / Nominal finite and positive
    bCntOk := (uPulseCount >= uMinPulses) AND (uPulseCount > 0); // 样本量达标且分母为正 / Sample count adequate, denominator positive
    IF NOT bNomOk THEN
        eState    := eFault;                          // 组态当量非法锁故障 / Illegal nominal latches fault
        uCodeLatch := 16#0003_00FA;                   // 码位：当量非法 / Code: illegal equivalent
        bError    := TRUE;                            // 故障级配对置位（R45）/ Fault flag paired
        uErrorId  := 16#0003_00FA;                    // 故障码回放 / Fault code replayed
    ELSIF NOT bVolOk THEN
        eState    := eFault;                          // 容积非法锁故障 / Illegal volume latches fault
        uCodeLatch := 16#0003_00F9;                   // 码位：容积非法 / Code: illegal volume
        bError    := TRUE;                            // 故障级配对置位 / Fault flag paired
        uErrorId  := 16#0003_00F9;                    // 故障码回放 / Fault code replayed
    ELSIF NOT bCntOk THEN
        eState    := eFault;                          // 样本不足锁故障 / Insufficient sample latches fault
        uCodeLatch := 16#0003_00F8;                   // 码位：样本不足 / Code: insufficient sample
        bError    := TRUE;                            // 故障级配对置位 / Fault flag paired
        uErrorId  := 16#0003_00F8;                    // 故障码回放 / Fault code replayed
    ELSE
        fMeasEquiv := fMeasuredMl / UDINT_TO_REAL(uPulseCount); // 实测当量，分母已验正 / Measured equivalent, denominator verified
        fDevPct := (fMeasEquiv - fNominalMlPerPulse) / fNominalMlPerPulse * DL_DPC_PCT; // 偏差百分数 / Deviation percent
        fNomAbs := ABS(fNominalMlPerPulse);           // 夹带基准幅值 / Clamp base magnitude
        fCorrEquiv := fNominalMlPerPulse * fNominalMlPerPulse / fMeasEquiv; // 反向修正：实测偏大则当量调小 / Inverse correction
        fCorrEquiv := MIN(MAX(fCorrEquiv, DL_DPC_LO * fNomAbs), DL_DPC_HI * fNomAbs); // 夹在组态 0.5~2.0 倍带内 / Clamp to 0.5..2.0x band
        fMeasuredMlPerPulse   := fMeasEquiv;          // 输出实测当量 / Emit measured equivalent
        fDeviationPct         := fDevPct;             // 输出偏差 / Emit deviation
        fCorrectedMlPerPulse  := fCorrEquiv;          // 输出修正当量 / Emit corrected equivalent
        bError    := FALSE;                           // 计算成功清故障 / Clear fault on success
        uCodeLatch := 16#0000_0000;                   // 清锁存码 / Clear latched code
        IF ABS(fDevPct) > fTolPct THEN
            uErrorId := 16#0003_00FB;                 // 告警级：偏差超限（不置 bError）/ Alarm: deviation out of band
        ELSE
            uErrorId := 16#0000_0000;                 // 无码 / No code
        END_IF
        eState := eDone;                              // 转完成态发单拍脉冲 / To done for one-scan pulse
        bBusy  := TRUE;                               // 计算当拍置忙（下拍由完成态清）/ Busy during compute scan
    END_IF
END_IF

// ---- 段 5｜故障态输出冻结回放（保持末次有效值，禁零值覆盖）----------------------
IF eState = eFault THEN
    bBusy    := FALSE;                                // 故障态清忙 / Clear busy in fault
    bDone    := FALSE;                                // 故障态不置完成 / Never done in fault
    bError   := TRUE;                                 // 故障标志保持 / Fault flag held
    uErrorId := uCodeLatch;                           // 故障码锁存回放 / Latched fault code replayed
END_IF

// ---- 段 6｜待机态默认清零（R27 输出保持语义：非保持量逐拍重算）------------------
IF eState = eIdle THEN
    bBusy  := FALSE;                                  // 待机清忙 / Idle clears busy
    bDone  := FALSE;                                  // 待机清完成脉冲 / Idle clears done pulse
    IF uErrorId = 16#0003_00F7 THEN
        uErrorId := 16#0000_0000;                     // 中止信息码单拍回落 / Abort info code single-scan fallback
    END_IF
END_IF
END_FUNCTION_BLOCK

(* ---- FB_DL_DustCollectorPulse.st ---- *)
(*
  ==================================================================
  组件名 Component  : FB_DL_DustCollectorPulse
  分类   Category   : DL_Device
  复杂度 Complexity  : 中
  版本   Version    : 1.0.0
  功能   Purpose    : 布袋除尘器脉冲反吹。压差分级触发（fDpStart 开 /
                      fDpStop 关回差）；轮巡脉阀（tPulse 得电 → tInterval 间
                      隔 → 下一阀）；清灰无效劣化报警：整轮巡完且压差仍高于
                      fDpHigh 累轮 nRoundMax 轮 → 锁存 bDpHighAlm。LBP 三段
                      骨架（命令→监视→判定）。
  来源   Source     : T2-2-lbp（LBP 三段骨架）
  溯源   Origin     : IEC 61131-3 标准语义的道莅防御性实现；压差回差与脉阀
                      轮巡为行业公知工程语义，clean-room 自研实现，未复制
                      LBP 或任何厂商私有库源码。
  平台   Platform   : 纯 IEC 61131-3（Standard.library: TON / R_TRIG，无私有库）
  分工声明 Split     : 与 FB_DL_SprayNozzleBank 分工——后者做喷嘴组搭接排
                      布，本件做除尘压差触发脉阀轮巡。
  作者   Author     : 道莅代码库 · PLC 编程专家（R59）
  ------------------------------------------------------------------
  边界 Boundary     :
                      一 安全语义：报警 / 非有限压差 / 停止时全阀输出统一出
                         口强制 FALSE（安全侧单点映射，R191）；
                      二 组态域闸：nValves ∈ [1..8]，越域锁存 bError（解除
                         = bReset 沿，R188）；
                      三 阀脉冲窗 / 间隔窗到期即迁（窗口末退出迁移，纪律④）；
                      四 非有限压差置 bBad（纪律②）挂起触发与判定不误报；
                      五 报警锁存解除路径 = bReset 沿（唯一路径，R188 声明）；
                      六 定时器与沿检测全部段 0 无条件周期刷新（R7）；
                      七 无全局变量、无外部变量声明、无物理地址寻址。
  修订记录 Revision  :
    2026-11-21  v1.0.0  R59 首版（批 3 · 序号 14）
  ==================================================================
*)

FUNCTION_BLOCK FB_DL_DustCollectorPulse
VAR_INPUT
    fDpKpa    : LREAL := 0.0;   // 除尘器压差反馈 [千帕] / the dust collector differential pressure [kilopascal]
    fDpStart  : LREAL := 1.2;   // 反吹启动压差阈值 [千帕] / the cleaning start threshold [kilopascal]
    fDpStop   : LREAL := 0.9;   // 反吹停止压差阈值（回差下限）[千帕] / the cleaning stop threshold [kilopascal]
    fDpHigh   : LREAL := 2.0;   // 清灰无效判定压差 [千帕] / the ineffective cleaning verdict pressure [kilopascal]
    nValves   : INT := 8;       // 脉阀数 [只]，域 1..8 / the valve count, one through eight
    tPulse    : TIME := T#150MS; // 脉阀得电时长 [毫秒] / the valve pulse duration [millisecond]
    tInterval : TIME := T#5S;   // 阀间间隔时长 [毫秒] / the valve interval [millisecond]
    nRoundMax : UDINT := 3;     // 无效判定累轮限 [轮] / the ineffective round bound
    bStop     : BOOL := FALSE;  // 停止指令，电平生效 [-] / the stop command, level effective
    bReset    : BOOL := FALSE;  // 报警与组态复位，上升沿生效 [-] / the alarm and config reset, rising edge
END_VAR
VAR_OUTPUT
    aValve     : ARRAY[0..7] OF BOOL; // 脉阀输出组 [-] / the valve outlets
    nValveIdx  : INT  := -1;  // 当前脉阀索引，-1 = 无 [只] / the current valve index, minus one when none
    bValveOn   : BOOL := FALSE; // 当前阀得电进行中 [-] / the current valve energized
    bCleaning  : BOOL := FALSE; // 反吹轮巡进行指示 [-] / the cleaning round robin indicator
    bDpHighAlm : BOOL := FALSE; // 清灰无效劣化报警锁存（解除 = bReset 沿）[-] / the ineffective cleaning alarm latch
    nRoundCnt  : UDINT := 0;  // 无效累轮计数 [轮] / the ineffective round count
    bBad       : BOOL := FALSE; // 非有限压差实时标志 [-] / the non finite pressure flag
    bError     : BOOL := FALSE; // 组态域闸故障锁存 [-] / the config gate fault latch
END_VAR
VAR CONSTANT
    DL_DCP_VMAX   : INT  := 8;           // 阀容量上界 [只] / the valve capacity bound
    DL_DCP_CNTMAX : UDINT := 4294967294; // 计数防回绕上界 [轮] / the counter anti wrap clamp bound
END_VAR
VAR
    _bRun    : BOOL := FALSE; // 轮巡运行锁存（压差回差驱动）/ the round robin run latch, driven by the hysteresis
    _nValve  : INT := 0;   // 轮巡阀寄存 [只] / the round robin valve register
    _bOn     : BOOL := FALSE; // 阀得电相位寄存 / the valve on phase register
    _bWrap   : BOOL := FALSE; // 整轮回绕捕获寄存 / the full round wrap capture register
    _bInit   : BOOL := FALSE; // 首拍初始化标志（R310，真实使用：首拍清阀输出）/ the first scan flag, real use
    _nI      : DINT;       // 阀遍历索引 / the valve loop index
    _bFinDp  : BOOL;       // 压差有限工作量 [-] / the pressure finiteness work flag
    rtReset  : R_TRIG;     // 复位沿，段 0 无条件刷新 / the reset edge
    tonPulse : TON;        // 阀脉冲窗，段 0 无条件刷新 / the valve pulse window
    tonGap   : TON;        // 阀间间隔窗，段 0 无条件刷新 / the valve interval window
END_VAR

// 段 0｜定时器与沿检测无条件周期刷新（禁入分支，R7）/ segment 0, the unconditional refresh
rtReset(CLK := bReset); // 复位沿 / the reset edge
tonPulse(IN := _bOn, PT := tPulse); // 阀脉冲窗 / the valve pulse window
tonGap(IN := _bRun AND (NOT _bOn) AND (NOT tonGap.Q), PT := tInterval); // 间隔窗（自复位单发，R188）/ the interval self reset window

// 段 1｜首拍初始化（R310 真实使用路径）：阀输出显式清零 / segment 1, the first scan init
IF NOT _bInit THEN // 首拍一拍 / the first scan
    _bInit := TRUE; // 置首拍标志 / raise the flag
    FOR _nI := 0 TO DL_DCP_VMAX - 1 DO // 全阀清零 / clear all the valves
        aValve[_nI] := FALSE; // 阀输出清零 / clear the valve outlet
    END_FOR
END_IF

// 段 2｜组态域闸与复位（边界二五，解除路径 = bReset 沿，R188）/ segment 2, the config gate and the reset
IF (nValves < 1) OR (nValves > DL_DCP_VMAX) THEN // 阀数越域 / the valve count out of domain
    bError := TRUE; // 置域闸锁存 / raise the config latch
END_IF
IF rtReset.Q THEN // 复位沿 / the reset edge
    bError := FALSE; // 清域闸锁存 / clear the config latch
    bDpHighAlm := FALSE; // 清劣化报警（唯一解除路径）/ clear the alarm
    nRoundCnt := 0; // 清累轮计数 / clear the round count
END_IF

// 段 3｜压差有限性与回差触发（边界四）/ segment 3, the pressure finiteness and the hysteresis
_bFinDp := (fDpKpa = fDpKpa) AND ((fDpKpa - fDpKpa) = (fDpKpa - fDpKpa)); // 压差有限双判据（R79）/ the finiteness dual verdicts
bBad := NOT _bFinDp; // 拒收实时标志（R191 名实双出口）/ the rejection flag
IF _bFinDp AND (NOT bError) THEN // 有效压差才参与触发 / only the valid pressure drives the trigger
    IF (NOT _bRun) AND (fDpKpa > fDpStart) THEN // 超启动阈值开轮巡 / beyond the start threshold, run
        _bRun := TRUE; // 开轮巡 / start the round robin
    ELSIF _bRun AND (fDpKpa < fDpStop) THEN // 低于回差下限停轮巡 / below the stop threshold, halt
        _bRun := FALSE; // 停轮巡 / halt
        _bOn := FALSE; // 阀断电 / drop the valve
        _nValve := 0; // 阀寄存归零 / reset the valve register
    END_IF
END_IF

// 段 4｜轮巡相位消化（阀脉冲窗与间隔窗窗口末退出迁移，边界三）/ segment 4, the round robin consume
IF _bOn THEN // 阀得电相位 / the valve on phase
    IF tonPulse.Q THEN // 脉冲窗到期（窗口末退出迁移）/ the pulse expired
        _bOn := FALSE; // 阀断电进间隔 / drop the valve into the interval
    END_IF
ELSIF _bRun AND (NOT bError) AND (NOT bDpHighAlm) AND (NOT bStop) AND _bFinDp THEN // 间隔相位（有效运行窗）/ the interval phase in the valid window
    IF tonGap.Q THEN // 间隔窗到期（自复位单发，窗口末退出迁移）/ the interval expired, self reset one shot
        _nValve := _nValve + 1; // 阀推进 / advance the valve
        IF _nValve >= nValves THEN // 整轮回绕 / the full round wrap
            _nValve := 0; // 回首阀 / back to the first valve
            _bWrap := TRUE; // 捕获整轮 / capture the full round
        END_IF
        _bOn := TRUE; // 下一阀得电 / energize the next valve
    END_IF
END_IF

// 段 5｜清灰无效劣化判定（整轮巡完且压差仍高，累轮达限锁存，边界五）/ segment 5, the ineffective cleaning verdict
IF _bWrap THEN // 整轮捕获沿 / the full round captured
    _bWrap := FALSE; // 捕获消化 / absorb the capture
    IF _bFinDp AND (fDpKpa > fDpHigh) THEN // 轮末压差仍高于判定限 / the pressure still high at the round end
        IF nRoundCnt < DL_DCP_CNTMAX THEN // 计数防回绕 / the wrap guard
            nRoundCnt := nRoundCnt + 1; // 累轮推进 / advance the round count
        END_IF
        IF nRoundCnt >= nRoundMax THEN // 达累轮限 / at the round bound
            bDpHighAlm := TRUE; // 置劣化报警锁存（成因独立，R190）/ raise the alarm latch
            _bRun := FALSE; // 停轮巡（报警安全侧）/ halt the round robin
            _bOn := FALSE; // 阀断电 / drop the valve
        END_IF
    END_IF
END_IF

// 段 6｜统一出口：阀输出单点安全映射（边界一）/ segment 6, the unified outlet
FOR _nI := 0 TO DL_DCP_VMAX - 1 DO // 全阀重映射 / remap all the valves
    aValve[_nI] := FALSE; // 先全断（安全侧基线）/ all off first, the safe baseline
END_FOR
IF _bOn AND (NOT bError) AND (NOT bDpHighAlm) AND (NOT bStop) AND _bFinDp THEN // 阀得电有效窗 / the valid energize window
    IF (_nValve >= 0) AND (_nValve < nValves) THEN // 阀界闸（防越界写）/ the valve bound gate
        aValve[_nValve] := TRUE; // 当前阀得电 / the current valve on
    END_IF
END_IF
nValveIdx := _nValve; // 阀索引出口 / the valve index outlet
bValveOn := _bOn; // 得电指示（R191 名实双出口）/ the energize indicator
bCleaning := _bRun; // 轮巡指示 / the round robin indicator
END_FUNCTION_BLOCK

(* ---- FB_DL_DustFreehoodPress.st ---- *)
(*==============================================================================
 * 组件名称 (Component)  : FB_DL_DustFreehoodPress
 * 溯源说明 (Provenance) : 道莅 clean-room 防御性实现（路线图 L363 已登记项）
 * 所属子库 (Sublibrary) : DL_Device / CleanroomDiag
 * 当前版本 (Version)    : 1.0.0
 * 兼容性   (Platform)   : CODESYS 3.5 / TwinCAT 3 / 汇川 InoProShop；
 *                         纯 IEC 61131-3（第 3 版），零标准库依赖
 * 组件分类 (Category)   : 功能块（FUNCTION_BLOCK）· 洁净风帽压差梯度监视
 * 功能一句话 (Summary)  : 多房间压差梯度校核 + 倒序最差相邻对定位 + 级联告警。
 * 边界与安全 (Boundary) : ①任一传感器失效 → 全列输出保持 + 告警（安全侧）；
 *                         ②房间数小于 2 → 配置非法码不判定；
 *                         ③压差非有限或负值 → 视同传感器失效（安全侧）；
 *                         ④相邻对下标全程钳位（禁越界访问）；
 *                         ⑤梯度约定：房间序号递增方向压差递减（洁净度梯度）。
 * 错误码    : 16#0003_0387 传感器失效（任一房间或通道失效）——故障级（持续态）
 *             16#0003_0388 级联梯度不足（最差相邻对低于门限）——故障级（持续态）
 *             16#0003_0389 配置非法（房间数不足 2）——故障级（持续态）
 * 码位总账  : 16#0003_0387 用 / 16#0003_0388 用 / 16#0003_0389 用
 * 修改记录  : v1.0.0 R26 初版
 *==============================================================================*)
FUNCTION_BLOCK FB_DL_DustFreehoodPress
VAR_INPUT
    afPress     : ARRAY[*] OF LREAL; // 各房间压差 [Pa]（序号递增为洁净度递增方向）/ Room differential pressures [Pa]
    fMinCascade : LREAL; // 相邻级最小梯度 [Pa] / Minimum adjacent cascade step [Pa]
    bSensorOk   : BOOL;  // 传感器通道自诊断 OK / Sensor channel self-check OK
END_VAR
VAR_OUTPUT
    bCascadeOk : BOOL; // 梯度全部达标 / All cascade steps qualified
    uWorstPair : UINT; // 倒序最差相邻对索引（压差[i]-压差[i+1] 最小者的 i）/ Worst adjacent pair index
    bRankAlarm : BOOL; // 级联排序告警 / Cascade ranking alarm
    eErr       : UDINT; // 本周期错误码，0=无错 / Error code this cycle, 0 = none
END_VAR
VAR
    iRooms  : INT;  // 房间数 / Room count
    i       : INT;  // 相邻对游标 / Adjacent pair cursor
    iWorst  : INT;  // 最差对内部值 / Worst pair internal
    fStep   : LREAL; // 当前相邻对梯度 / Current adjacent step
    fWorst  : LREAL; // 最差梯度值 / Worst gradient value
    bHold   : BOOL;  // 保持态判据 / Hold-state predicate
    fGrd    : LREAL; // 压差守卫副本 / Pressure guard copy
END_VAR

// ---------- 周期起点：错误码先清（持续态随后重置） ----------
eErr := 0;

// ---------- 配置防御：房间数不足 2 不判定 ----------
iRooms := UPPER_BOUND(afPress, 1) + 1;        // 房间数 / Room count
IF iRooms < 2 THEN
    bCascadeOk := FALSE;                      // 不判定安全侧 / Safe-side default
    uWorstPair := 0;                          // 索引缺省 / Index default
    bRankAlarm := FALSE;
    eErr := 16#0003_0389;                     // 配置非法码 / Illegal configuration code
    RETURN;
END_IF

// ---------- 传感器失效防御：全列保持（安全侧） ----------
bHold := (NOT bSensorOk) OR (fMinCascade <= 0.0) OR (fMinCascade <> fMinCascade);
IF bHold THEN
    IF NOT bSensorOk THEN
        bRankAlarm := TRUE;                   // 失效告警 / Failure alarm
        eErr := 16#0003_0387;                 // 传感器失效码 / Sensor failure code
    ELSE
        eErr := 16#0003_0389;                 // 门限非法视同配置非法 / Illegal threshold as config fault
    END_IF
    // bCascadeOk 与 uWorstPair 保持上拍锁存值（禁清零防误放行）/ Outputs held, no clear
    RETURN;
END_IF

// ---------- 逐相邻对校核：梯度递减约定（下标钳位） ----------
bCascadeOk := TRUE;                           // 先假设全达标 / Assume all qualified
iWorst := 0;
fWorst := 1.0E30;                             // 哨兵极大值 / Sentinel huge
FOR i := 0 TO iRooms - 2 DO
    fGrd := afPress[i];                       // 上游房间压差 / Upstream pressure
    IF (fGrd <> fGrd) OR ((fGrd - fGrd) <> (fGrd - fGrd)) OR (fGrd < 0.0) THEN
        bHold := TRUE;                        // 非有限或负值视同失效 / Non-finite or negative as failure
        eErr := 16#0003_0387;                 // 传感器失效码 / Sensor failure code
    ELSE
        fStep := afPress[i] - afPress[i + 1]; // 相邻对梯度 / Adjacent step
        IF fStep < fWorst THEN
            fWorst := fStep;                  // 更新最差值 / Update worst value
            iWorst := i;                      // 更新最差对索引 / Update worst index
        END_IF
        IF fStep < fMinCascade THEN
            bCascadeOk := FALSE;              // 梯度不足 / Step below threshold
        END_IF
    END_IF
END_FOR

// ---------- 失效保持出口：输出锁存不清（防误放行） ----------
IF bHold THEN
    bRankAlarm := TRUE;                       // 保持态告警 / Hold-state alarm
    RETURN;                                   // bCascadeOk/uWorstPair 锁存 / Outputs latched
END_IF

// ---------- 结论输出：最差对索引与告警 ----------
uWorstPair := INT_TO_UINT(iWorst);            // 倒序最差对索引 / Worst pair index exposed
IF bCascadeOk THEN
    bRankAlarm := FALSE;                      // 全达标不告警 / No alarm when qualified
ELSE
    bRankAlarm := TRUE;                       // 梯度不足告警 / Under-threshold alarm
    eErr := 16#0003_0388;                     // 级联梯度不足码 / Cascade deficit code
END_IF

END_FUNCTION_BLOCK
